(* IEC 61131-3 sources: rusty/tests/lit/single/conversion, 25 files *)

(* ---- to_string_unsupported.st ---- *)
// RUN: not %COMPILE %s 2>&1 | %CHECK %s
// A type with no TO_STRING monomorphization must not silently mis-dispatch to TO_STRING__STRING
// (which reinterprets the argument's bytes and crashes at runtime). Instead the missing
// monomorphization is materialized as an external declaration and surfaces as a link-time undefined
// symbol — a clean, uniform failure for scalar and aggregate returns alike. A user STRUCT never gets
// a monomorph, so this stays valid as follow-up PRs add the remaining scalar conversions.
TYPE MyStruct : STRUCT x : DINT; END_STRUCT END_TYPE

FUNCTION main : DINT
VAR
    st : MyStruct;
    s : STRING;
END_VAR
    // CHECK: {{.*}}TO_STRING__MyStruct{{.*}}
    s := TO_STRING(st);
END_FUNCTION

(* ---- bit_to_real.st ---- *)
// RUN: %COMPILE %s && %RUN | %CHECK %s
//
// BOOL and the bit string types widen to REAL and LREAL by value. BOOL, BYTE and WORD fit a REAL
// exactly, and DWORD fits an LREAL exactly. A REAL keeps 24 bits of mantissa, so a DWORD or LWORD
// above 2^24 is rounded to the nearest representable value on the way in, without a diagnostic.
// These conversions have the named form only; the generic TO_REAL and TO_LREAL take numeric sources.

FUNCTION main
VAR
    umax : LWORD := 0;
END_VAR
umax := umax - 1;   // 2^64 - 1

// BOOL
printf('%.1f %.1f %.1f %.1f$N', BOOL_TO_REAL(FALSE), BOOL_TO_REAL(TRUE), BOOL_TO_LREAL(FALSE), BOOL_TO_LREAL(TRUE));  // CHECK: 0.0 1.0 0.0 1.0

// BYTE and WORD, exact over the whole range
printf('%.0f %.0f %.0f %.0f$N', BYTE_TO_REAL(BYTE#255), BYTE_TO_LREAL(BYTE#255), WORD_TO_REAL(WORD#65535), WORD_TO_LREAL(WORD#65535));  // CHECK: 255 255 65535 65535

// DWORD: exact into LREAL, rounded into REAL above 2^24
printf('%.0f %.0f$N', DWORD_TO_LREAL(DWORD#16777217), DWORD_TO_LREAL(DWORD#4294967295));  // CHECK: 16777217 4294967295
printf('%.0f %.0f$N', DWORD_TO_REAL(DWORD#16777216),  DWORD_TO_REAL(DWORD#16777217));     // CHECK: 16777216 16777216
printf('%.0f$N',      DWORD_TO_REAL(DWORD#4294967295));                                   // CHECK: 4294967296

// LWORD into REAL: 2^24 is the last exact integer
printf('%.0f %.0f$N', LWORD_TO_REAL(LWORD#16777216), LWORD_TO_REAL(LWORD#16777217));          // CHECK: 16777216 16777216
printf('%.0f %.0f$N', LWORD_TO_REAL(LWORD#4294967296), LWORD_TO_REAL(LWORD#9007199254740993));  // CHECK: 4294967296 9007199254740992
printf('%.0f$N',      LWORD_TO_REAL(umax));                                                    // CHECK: 18446744073709551616

// LWORD into LREAL: 2^53 is the last exact integer
printf('%.0f %.0f$N', LWORD_TO_LREAL(LWORD#4611686018427387904), LWORD_TO_LREAL(LWORD#9007199254740993));  // CHECK: 4611686018427387904 9007199254740992
END_FUNCTION

(* ---- num_to_bool.st ---- *)
// RUN: %COMPILE %s && %RUN | %CHECK %s
//
// Every *_TO_BOOL conversion is FALSE for exactly zero and TRUE for everything else. It is not a
// lowest-bit test, a fraction is not truncated first, there is no epsilon, and NaN and the
// infinities are TRUE.

FUNCTION main
VAR
    umax : ULINT := 0;
    ninf : REAL;
END_VAR
umax := umax - 1;   // 2^64 - 1
ninf := -INF_REAL;

// signed integers
printf('%d %d %d %d %d$N', SINT_TO_BOOL(SINT#-128), SINT_TO_BOOL(SINT#0), INT_TO_BOOL(INT#2), INT_TO_BOOL(INT#256), INT_TO_BOOL(INT#-1));  // CHECK: 1 0 1 1 1
printf('%d %d %d %d$N',    INT_TO_BOOL(INT#0), INT_TO_BOOL(INT#1), DINT_TO_BOOL(DINT#65536), LINT_TO_BOOL(LINT#4294967296));                  // CHECK: 0 1 1 1

// unsigned integers
printf('%d %d %d %d$N', USINT_TO_BOOL(USINT#255), USINT_TO_BOOL(USINT#0), UINT_TO_BOOL(UINT#256), UDINT_TO_BOOL(UDINT#4294967295));  // CHECK: 1 0 1 1
printf('%d %d %d %d$N', USINT_TO_BOOL(USINT#1), UINT_TO_BOOL(UINT#0), UINT_TO_BOOL(UINT#65535), UDINT_TO_BOOL(UDINT#65536));         // CHECK: 1 0 1 1
printf('%d %d %d %d$N', ULINT_TO_BOOL(umax), ULINT_TO_BOOL(ULINT#9223372036854775807), ULINT_TO_BOOL(ULINT#4294967296), ULINT_TO_BOOL(ULINT#0));  // CHECK: 1 1 1 0

// reals
printf('%d %d %d %d$N', REAL_TO_BOOL(REAL#0.5), REAL_TO_BOOL(REAL#1.0E-30), REAL_TO_BOOL(REAL#0.0), REAL_TO_BOOL(-REAL#0.0));  // CHECK: 1 1 0 0
printf('%d %d %d$N',    REAL_TO_BOOL(NAN_REAL), REAL_TO_BOOL(INF_REAL), REAL_TO_BOOL(ninf));                                    // CHECK: 1 1 1
printf('%d %d %d$N',    LREAL_TO_BOOL(LREAL#-0.5), LREAL_TO_BOOL(LREAL#0.0), LREAL_TO_BOOL(NAN_LREAL));                          // CHECK: 1 0 1
printf('%d %d %d$N',    LREAL_TO_BOOL(LREAL#0.5), LREAL_TO_BOOL(-LREAL#0.0), LREAL_TO_BOOL(LREAL#1.0E-300));                     // CHECK: 1 0 1

// bit strings, a set bit above bit 0 is TRUE as well
printf('%d %d %d %d %d$N', BYTE_TO_BOOL(BYTE#2), BYTE_TO_BOOL(BYTE#0), WORD_TO_BOOL(WORD#256), DWORD_TO_BOOL(DWORD#65536), LWORD_TO_BOOL(LWORD#4294967296));  // CHECK: 1 0 1 1 1

// the generic form calls the named one
printf('%d %d %d %d$N', TO_BOOL(INT#256), TO_BOOL(REAL#0.5), TO_BOOL(ULINT#4294967296), TO_BOOL(BYTE#2));  // CHECK: 1 1 1 1
END_FUNCTION

(* ---- real_to_bit.st ---- *)
// RUN: %COMPILE %s && %RUN | %CHECK %s
//
// REAL and LREAL to the bit string types round half away from zero, then keep the low bits of the
// target width, so an out-of-range value wraps and a negative value lands at the top of the range.
// The rounded value first becomes a signed 64-bit integer; NaN, the infinities and anything outside
// that range become 2^63 instead, so BYTE, WORD and DWORD see 0 for them. LWORD is the exception:
// a value in [2^63, 2^64) converts exactly, and only NaN, the infinities, values below -2^63 and
// values at or above 2^64 give 2^63. Every cell was measured on CODESYS 3.5 SP22.
FUNCTION main
VAR
    ninf    : REAL;
    lninf   : LREAL;
    band_lo : LREAL := 9223372036854775808.0;   (* 2^63, the smallest LREAL above it is added below *)
    two64   : LREAL := 9223372036854775808.0;
END_VAR
ninf    := -INF_REAL;
lninf   := -INF_LREAL;
band_lo := band_lo + 2048.0;
two64   := two64 * 2.0;

// ---- REAL source: BYTE WORD DWORD LWORD
// rounding, ties away from zero
printf('%d %d %u %llu$N', REAL_TO_BYTE(REAL#0.4),  REAL_TO_WORD(REAL#0.4),  REAL_TO_DWORD(REAL#0.4),  REAL_TO_LWORD(REAL#0.4));   // CHECK: 0 0 0 0
printf('%d %d %u %llu$N', REAL_TO_BYTE(REAL#0.5),  REAL_TO_WORD(REAL#0.5),  REAL_TO_DWORD(REAL#0.5),  REAL_TO_LWORD(REAL#0.5));   // CHECK: 1 1 1 1
printf('%d %d %u %llu$N', REAL_TO_BYTE(REAL#0.6),  REAL_TO_WORD(REAL#0.6),  REAL_TO_DWORD(REAL#0.6),  REAL_TO_LWORD(REAL#0.6));   // CHECK: 1 1 1 1
printf('%d %d %u %llu$N', REAL_TO_BYTE(REAL#1.5),  REAL_TO_WORD(REAL#1.5),  REAL_TO_DWORD(REAL#1.5),  REAL_TO_LWORD(REAL#1.5));   // CHECK: 2 2 2 2
printf('%d %d %u %llu$N', REAL_TO_BYTE(REAL#2.5),  REAL_TO_WORD(REAL#2.5),  REAL_TO_DWORD(REAL#2.5),  REAL_TO_LWORD(REAL#2.5));   // CHECK: 3 3 3 3
printf('%d %d %u %llu$N', REAL_TO_BYTE(REAL#3.5),  REAL_TO_WORD(REAL#3.5),  REAL_TO_DWORD(REAL#3.5),  REAL_TO_LWORD(REAL#3.5));   // CHECK: 4 4 4 4
printf('%d %d %u %llu$N', REAL_TO_BYTE(REAL#-0.5), REAL_TO_WORD(REAL#-0.5), REAL_TO_DWORD(REAL#-0.5), REAL_TO_LWORD(REAL#-0.5));  // CHECK: 255 65535 4294967295 18446744073709551615
printf('%d %d %u %llu$N', REAL_TO_BYTE(REAL#-1.5), REAL_TO_WORD(REAL#-1.5), REAL_TO_DWORD(REAL#-1.5), REAL_TO_LWORD(REAL#-1.5));  // CHECK: 254 65534 4294967294 18446744073709551614
printf('%d %d %u %llu$N', REAL_TO_BYTE(REAL#-2.5), REAL_TO_WORD(REAL#-2.5), REAL_TO_DWORD(REAL#-2.5), REAL_TO_LWORD(REAL#-2.5));  // CHECK: 253 65533 4294967293 18446744073709551613
// range, wraps modulo the target width
printf('%d %d %u %llu$N', REAL_TO_BYTE(REAL#255.5),   REAL_TO_WORD(REAL#255.5),   REAL_TO_DWORD(REAL#255.5),   REAL_TO_LWORD(REAL#255.5));    // CHECK: 0 256 256 256
printf('%d %d %u %llu$N', REAL_TO_BYTE(REAL#256.0),   REAL_TO_WORD(REAL#256.0),   REAL_TO_DWORD(REAL#256.0),   REAL_TO_LWORD(REAL#256.0));    // CHECK: 0 256 256 256
printf('%d %d %u %llu$N', REAL_TO_BYTE(REAL#300.0),   REAL_TO_WORD(REAL#300.0),   REAL_TO_DWORD(REAL#300.0),   REAL_TO_LWORD(REAL#300.0));    // CHECK: 44 300 300 300
printf('%d %d %u %llu$N', REAL_TO_BYTE(REAL#-1.0),    REAL_TO_WORD(REAL#-1.0),    REAL_TO_DWORD(REAL#-1.0),    REAL_TO_LWORD(REAL#-1.0));     // CHECK: 255 65535 4294967295 18446744073709551615
printf('%d %d %u %llu$N', REAL_TO_BYTE(REAL#65536.0), REAL_TO_WORD(REAL#65536.0), REAL_TO_DWORD(REAL#65536.0), REAL_TO_LWORD(REAL#65536.0));  // CHECK: 0 0 65536 65536
printf('%d %d %u %llu$N', REAL_TO_BYTE(REAL#1.0E10),  REAL_TO_WORD(REAL#1.0E10),  REAL_TO_DWORD(REAL#1.0E10),  REAL_TO_LWORD(REAL#1.0E10));   // CHECK: 0 58368 1410065408 10000000000
printf('%d %d %u %llu$N', REAL_TO_BYTE(REAL#1.0E20),  REAL_TO_WORD(REAL#1.0E20),  REAL_TO_DWORD(REAL#1.0E20),  REAL_TO_LWORD(REAL#1.0E20));   // CHECK: 0 0 0 9223372036854775808
// not a number
printf('%d %d %u %llu$N', REAL_TO_BYTE(INF_REAL), REAL_TO_WORD(INF_REAL), REAL_TO_DWORD(INF_REAL), REAL_TO_LWORD(INF_REAL));  // CHECK: 0 0 0 9223372036854775808
printf('%d %d %u %llu$N', REAL_TO_BYTE(ninf),     REAL_TO_WORD(ninf),     REAL_TO_DWORD(ninf),     REAL_TO_LWORD(ninf));      // CHECK: 0 0 0 9223372036854775808
printf('%d %d %u %llu$N', REAL_TO_BYTE(NAN_REAL), REAL_TO_WORD(NAN_REAL), REAL_TO_DWORD(NAN_REAL), REAL_TO_LWORD(NAN_REAL));  // CHECK: 0 0 0 9223372036854775808

// ---- LREAL source: BYTE WORD DWORD LWORD
printf('%d %d %u %llu$N', LREAL_TO_BYTE(LREAL#0.5),     LREAL_TO_WORD(LREAL#0.5),     LREAL_TO_DWORD(LREAL#0.5),     LREAL_TO_LWORD(LREAL#0.5));      // CHECK: 1 1 1 1
printf('%d %d %u %llu$N', LREAL_TO_BYTE(LREAL#2.5),     LREAL_TO_WORD(LREAL#2.5),     LREAL_TO_DWORD(LREAL#2.5),     LREAL_TO_LWORD(LREAL#2.5));      // CHECK: 3 3 3 3
printf('%d %d %u %llu$N', LREAL_TO_BYTE(LREAL#-0.5),    LREAL_TO_WORD(LREAL#-0.5),    LREAL_TO_DWORD(LREAL#-0.5),    LREAL_TO_LWORD(LREAL#-0.5));     // CHECK: 255 65535 4294967295 18446744073709551615
printf('%d %d %u %llu$N', LREAL_TO_BYTE(LREAL#-2.5),    LREAL_TO_WORD(LREAL#-2.5),    LREAL_TO_DWORD(LREAL#-2.5),    LREAL_TO_LWORD(LREAL#-2.5));     // CHECK: 253 65533 4294967293 18446744073709551613
printf('%d %d %u %llu$N', LREAL_TO_BYTE(LREAL#255.5),   LREAL_TO_WORD(LREAL#255.5),   LREAL_TO_DWORD(LREAL#255.5),   LREAL_TO_LWORD(LREAL#255.5));    // CHECK: 0 256 256 256
printf('%d %d %u %llu$N', LREAL_TO_BYTE(LREAL#300.0),   LREAL_TO_WORD(LREAL#300.0),   LREAL_TO_DWORD(LREAL#300.0),   LREAL_TO_LWORD(LREAL#300.0));    // CHECK: 44 300 300 300
printf('%d %d %u %llu$N', LREAL_TO_BYTE(LREAL#-1.0),    LREAL_TO_WORD(LREAL#-1.0),    LREAL_TO_DWORD(LREAL#-1.0),    LREAL_TO_LWORD(LREAL#-1.0));     // CHECK: 255 65535 4294967295 18446744073709551615
printf('%d %d %u %llu$N', LREAL_TO_BYTE(LREAL#65536.0), LREAL_TO_WORD(LREAL#65536.0), LREAL_TO_DWORD(LREAL#65536.0), LREAL_TO_LWORD(LREAL#65536.0));  // CHECK: 0 0 65536 65536
printf('%d %d %u %llu$N', LREAL_TO_BYTE(LREAL#1.0E10),  LREAL_TO_WORD(LREAL#1.0E10),  LREAL_TO_DWORD(LREAL#1.0E10),  LREAL_TO_LWORD(LREAL#1.0E10));   // CHECK: 0 58368 1410065408 10000000000
printf('%d %d %u %llu$N', LREAL_TO_BYTE(LREAL#1.0E20),  LREAL_TO_WORD(LREAL#1.0E20),  LREAL_TO_DWORD(LREAL#1.0E20),  LREAL_TO_LWORD(LREAL#1.0E20));   // CHECK: 0 0 0 9223372036854775808
printf('%d %d %u %llu$N', LREAL_TO_BYTE(INF_LREAL), LREAL_TO_WORD(INF_LREAL), LREAL_TO_DWORD(INF_LREAL), LREAL_TO_LWORD(INF_LREAL));  // CHECK: 0 0 0 9223372036854775808
printf('%d %d %u %llu$N', LREAL_TO_BYTE(lninf),     LREAL_TO_WORD(lninf),     LREAL_TO_DWORD(lninf),     LREAL_TO_LWORD(lninf));      // CHECK: 0 0 0 9223372036854775808
printf('%d %d %u %llu$N', LREAL_TO_BYTE(NAN_LREAL), LREAL_TO_WORD(NAN_LREAL), LREAL_TO_DWORD(NAN_LREAL), LREAL_TO_LWORD(NAN_LREAL));  // CHECK: 0 0 0 9223372036854775808

// ---- the 64-bit band: LWORD keeps [2^63, 2^64) exact, the narrower targets go through the signed path
printf('%u %llu$N', LREAL_TO_DWORD(LREAL#1.0E19), LREAL_TO_LWORD(LREAL#1.0E19));   // CHECK: 0 10000000000000000000
printf('%llu %llu$N', LREAL_TO_LWORD(band_lo), LREAL_TO_LWORD(LREAL#1.8E19));      // CHECK: 9223372036854777856 18000000000000000000
printf('%llu %llu$N', LREAL_TO_LWORD(two64), LREAL_TO_LWORD(LREAL#-1.0E19));       // CHECK: 9223372036854775808 9223372036854775808
printf('%llu$N', REAL_TO_LWORD(REAL#1.0E19));                                       // CHECK: 9999999980506447872

// ---- the generic form calls the named one
printf('%d %d %u %llu$N', TO_BYTE(REAL#300.0), TO_WORD(LREAL#-1.0), TO_DWORD(REAL#1.0E10), TO_LWORD(LREAL#-0.5));  // CHECK: 44 65535 1410065408 18446744073709551615
END_FUNCTION

(* ---- real_trunc_int.st ---- *)
// RUN: %COMPILE %s && %RUN | %CHECK %s
FUNCTION main
    printf('%d$N', REAL_TRUNC_SINT(5.6));       // CHECK: 5
    printf('%d$N', REAL_TRUNC_USINT(5.6));      // CHECK: 5
    printf('%d$N', REAL_TRUNC_INT(5.6));        // CHECK: 5
    printf('%d$N', REAL_TRUNC_UINT(5.6));       // CHECK: 5
    printf('%d$N', REAL_TRUNC_INT(5.6));        // CHECK: 5
    printf('%d$N', REAL_TRUNC_UINT(5.6));       // CHECK: 5
    printf('%d$N', REAL_TRUNC_DINT(5.6));       // CHECK: 5
    printf('%d$N', REAL_TRUNC_UDINT(5.6));      // CHECK: 5
    printf('%d$N', REAL_TRUNC_LINT(5.6));       // CHECK: 5
    printf('%d$N', REAL_TRUNC_ULINT(5.6));      // CHECK: 5

    printf('%d$N', REAL_TRUNC_SINT(-5.6));      // CHECK: -5
    printf('%d$N', REAL_TRUNC_INT(-5.6));       // CHECK: -5
    printf('%d$N', REAL_TRUNC_DINT(-5.6));      // CHECK: -5
    printf('%d$N', REAL_TRUNC_LINT(-5.6));      // CHECK: -5
END_FUNCTION

(* ---- string_to_based_literals.st ---- *)
// STRING_TO integer and bit-string conversions accept IEC based literals and nothing else.
// RUN: %COMPILE %s && %RUN | %CHECK %s

FUNCTION main
    printf('byte_hex=%d$N', STRING_TO_BYTE('16#FF'));        // CHECK: byte_hex=255
    printf('word_octal=%d$N', STRING_TO_WORD('8#777'));      // CHECK-NEXT: word_octal=511
    printf('dword_binary=%d$N', STRING_TO_DWORD('2#1010'));  // CHECK-NEXT: dword_binary=10
    printf('dint_binary=%d$N', STRING_TO_DINT('2#1010'));    // CHECK-NEXT: dint_binary=10
    printf('lint_binary=%d$N', STRING_TO_LINT('2#1010'));    // CHECK-NEXT: lint_binary=10
    printf('lword_lower_hex=%d$N', STRING_TO_LWORD('16#ff'));// CHECK-NEXT: lword_lower_hex=255
    printf('dint_hex=%d$N', STRING_TO_DINT('16#FF'));        // CHECK-NEXT: dint_hex=255
    printf('lint_hex=%d$N', STRING_TO_LINT('16#FF'));        // CHECK-NEXT: lint_hex=255
    printf('dint_octal=%d$N', STRING_TO_DINT('8#77'));       // CHECK-NEXT: dint_octal=63
    printf('lint_octal=%d$N', STRING_TO_LINT('8#77'));       // CHECK-NEXT: lint_octal=63
    printf('udint_grouped_hex=%d$N', STRING_TO_UDINT('16#FF_FF')); // CHECK-NEXT: udint_grouped_hex=65535
    printf('ulint_trimmed_hex=%d$N', STRING_TO_ULINT(' 16#FF ')); // CHECK-NEXT: ulint_trimmed_hex=255
    printf('missing_digits=%d$N', STRING_TO_UDINT('16#'));   // CHECK-NEXT: missing_digits=0
    printf('invalid_digit=%d$N', STRING_TO_UDINT('16#GG'));  // CHECK-NEXT: invalid_digit=0
    printf('unsupported_radix=%d$N', STRING_TO_UDINT('10#42')); // CHECK-NEXT: unsupported_radix=0
    printf('signed_hex=%d$N', STRING_TO_UDINT('+16#FF'));    // CHECK-NEXT: signed_hex=0

    // Based literals are unsigned; a sign on either side of the radix is rejected.
    printf('negative_hex=%d$N', STRING_TO_DINT('-16#FF'));   // CHECK-NEXT: negative_hex=0
    printf('hex_negative=%d$N', STRING_TO_DINT('16#-FF'));   // CHECK-NEXT: hex_negative=0
    printf('binary_negative=%d$N', STRING_TO_SINT('2#-1'));  // CHECK-NEXT: binary_negative=0

    // Underscores group digits; they may not lead, trail or double up.
    printf('leading_underscore=%d$N', STRING_TO_UDINT('16#_FF'));  // CHECK-NEXT: leading_underscore=0
    printf('trailing_underscore=%d$N', STRING_TO_UDINT('16#FF_')); // CHECK-NEXT: trailing_underscore=0
    printf('double_underscore=%d$N', STRING_TO_UDINT('16#F__F')); // CHECK-NEXT: double_underscore=0
    printf('decimal_grouped=%d$N', STRING_TO_UDINT('1_000'));     // CHECK-NEXT: decimal_grouped=1000
    printf('decimal_leading_us=%d$N', STRING_TO_UDINT('_1'));     // CHECK-NEXT: decimal_leading_us=0
    printf('decimal_double_us=%d$N', STRING_TO_UDINT('1__0'));    // CHECK-NEXT: decimal_double_us=0

    // C-style radix prefixes are not Structured Text literals.
    printf('byte_c_binary=%d$N', STRING_TO_BYTE('0b1010'));   // CHECK-NEXT: byte_c_binary=0
    printf('lword_c_binary=%d$N', STRING_TO_LWORD('0B1010')); // CHECK-NEXT: lword_c_binary=0
    printf('dint_c_hex=%d$N', STRING_TO_DINT('0x7F'));        // CHECK-NEXT: dint_c_hex=0
    printf('ulint_c_hex=%d$N', STRING_TO_ULINT('0X7F'));      // CHECK-NEXT: ulint_c_hex=0

    // A hexadecimal bit pattern that does not fit the signed target is rejected, not reinterpreted.
    printf('int_hex_max=%d$N', STRING_TO_INT('16#7FFF'));          // CHECK-NEXT: int_hex_max=32767
    printf('int_hex_all_ones=%d$N', STRING_TO_INT('16#FFFF'));     // CHECK-NEXT: int_hex_all_ones=0
    printf('word_hex_all_ones=%d$N', STRING_TO_WORD('16#FFFF'));   // CHECK-NEXT: word_hex_all_ones=65535
END_FUNCTION

(* ---- string_to_bool.st ---- *)
// STRING_TO_BOOL accepts true values and rejects malformed values.
// RUN: %COMPILE %s && %RUN | %CHECK %s

FUNCTION main
    printf('garbage=%d$N', STRING_TO_BOOL('garbage'));       // CHECK: garbage=0
    printf('numeric_one=%d$N', STRING_TO_BOOL('1'));         // CHECK-NEXT: numeric_one=1
    printf('upper_true=%d$N', STRING_TO_BOOL('TRUE'));       // CHECK-NEXT: upper_true=1
    printf('lower_true=%d$N', STRING_TO_BOOL('true'));       // CHECK-NEXT: lower_true=1
    printf('trimmed_true=%d$N', STRING_TO_BOOL('  true  ')); // CHECK-NEXT: trimmed_true=1
    printf('numeric_zero=%d$N', STRING_TO_BOOL('0'));        // CHECK-NEXT: numeric_zero=0
    printf('numeric_two=%d$N', STRING_TO_BOOL('2'));         // CHECK-NEXT: numeric_two=0
    printf('false=%d$N', STRING_TO_BOOL('false'));           // CHECK-NEXT: false=0
    printf('suffix=%d$N', STRING_TO_BOOL('TRUEX'));          // CHECK-NEXT: suffix=0
END_FUNCTION

(* ---- string_to_calendar.st ---- *)
// STRING_TO_DATE, STRING_TO_DT, and STRING_TO_TOD accept exactly the calendar literals of their type.
// RUN: %COMPILE %s && %RUN | %CHECK %s

FUNCTION main
    // Valid prefixed literals parse for each target type.
    printf('date_valid=%s$N', REF(DATE_TO_STRING(STRING_TO_DATE('D#2024-02-29')))); // CHECK: date_valid=D#2024-02-29
    printf('dt_valid=%s$N', REF(DT_TO_STRING(STRING_TO_DT('DT#2024-01-01-12:00:00')))); // CHECK-NEXT: dt_valid=DT#2024-01-01-12:00:00
    printf('tod_valid=%s$N', REF(TOD_TO_STRING(STRING_TO_TOD('TOD#12:00:00')))); // CHECK-NEXT: tod_valid=TOD#12:00:00

    // Empty input returns each type's zero value.
    printf('date_empty=%s$N', REF(DATE_TO_STRING(STRING_TO_DATE('')))); // CHECK-NEXT: date_empty=D#1970-01-01
    printf('dt_empty=%s$N', REF(DT_TO_STRING(STRING_TO_DT('')))); // CHECK-NEXT: dt_empty=DT#1970-01-01-00:00:00
    printf('tod_empty=%s$N', REF(TOD_TO_STRING(STRING_TO_TOD('')))); // CHECK-NEXT: tod_empty=TOD#00:00:00

    // Malformed input returns each type's zero value.
    printf('date_garbage=%s$N', REF(DATE_TO_STRING(STRING_TO_DATE('not a date')))); // CHECK-NEXT: date_garbage=D#1970-01-01
    printf('dt_garbage=%s$N', REF(DT_TO_STRING(STRING_TO_DT('$00')))); // CHECK-NEXT: dt_garbage=DT#1970-01-01-00:00:00
    printf('tod_garbage=%s$N', REF(TOD_TO_STRING(STRING_TO_TOD('bad')))); // CHECK-NEXT: tod_garbage=TOD#00:00:00

    // Each conversion rejects a literal prefix for a different calendar type.
    printf('date_wrong_prefix=%s$N', REF(DATE_TO_STRING(STRING_TO_DATE('TOD#12:45:00')))); // CHECK-NEXT: date_wrong_prefix=D#1970-01-01
    printf('dt_wrong_prefix=%s$N', REF(DT_TO_STRING(STRING_TO_DT('D#2024-01-01')))); // CHECK-NEXT: dt_wrong_prefix=DT#1970-01-01-00:00:00
    printf('tod_wrong_prefix=%s$N', REF(TOD_TO_STRING(STRING_TO_TOD('DT#2024-01-01-12:00:00')))); // CHECK-NEXT: tod_wrong_prefix=TOD#00:00:00

    // Out-of-range date and time fields are rejected.
    printf('date_invalid_day=%s$N', REF(DATE_TO_STRING(STRING_TO_DATE('D#2024-02-30')))); // CHECK-NEXT: date_invalid_day=D#1970-01-01
    printf('dt_invalid_hour=%s$N', REF(DT_TO_STRING(STRING_TO_DT('DT#2024-01-01-25:00:00')))); // CHECK-NEXT: dt_invalid_hour=DT#1970-01-01-00:00:00
    printf('tod_invalid_minute=%s$N', REF(TOD_TO_STRING(STRING_TO_TOD('TOD#12:60:00')))); // CHECK-NEXT: tod_invalid_minute=TOD#00:00:00

    // Values outside the representable range return the zero value.
    printf('date_low_range=%s$N', REF(DATE_TO_STRING(STRING_TO_DATE('D#1969-12-31')))); // CHECK-NEXT: date_low_range=D#1970-01-01
    printf('dt_low_range=%s$N', REF(DT_TO_STRING(STRING_TO_DT('DT#1969-12-31-23:59:59')))); // CHECK-NEXT: dt_low_range=DT#1970-01-01-00:00:00
    printf('tod_high_range=%s$N', REF(TOD_TO_STRING(STRING_TO_TOD('TOD#25:00:00')))); // CHECK-NEXT: tod_high_range=TOD#00:00:00
    printf('date_high_range=%s$N', REF(DATE_TO_STRING(STRING_TO_DATE('D#2106-02-08')))); // CHECK-NEXT: date_high_range=D#1970-01-01
    printf('dt_high_range=%s$N', REF(DT_TO_STRING(STRING_TO_DT('DT#2106-02-08-00:00:00')))); // CHECK-NEXT: dt_high_range=DT#1970-01-01-00:00:00
    printf('tod_low_range=%s$N', REF(TOD_TO_STRING(STRING_TO_TOD('TOD#-1:00:00')))); // CHECK-NEXT: tod_low_range=TOD#00:00:00

    // DATE rejects fractions, DT drops them, and TOD preserves milliseconds.
    printf('date_fraction=%s$N', REF(DATE_TO_STRING(STRING_TO_DATE('D#2024-01-01.500')))); // CHECK-NEXT: date_fraction=D#1970-01-01
    printf('dt_fraction=%s$N', REF(DT_TO_STRING(STRING_TO_DT('DT#2024-01-01-12:00:00.500')))); // CHECK-NEXT: dt_fraction=DT#2024-01-01-12:00:00
    printf('tod_fraction=%s$N', REF(TOD_TO_STRING(STRING_TO_TOD('TOD#12:00:00.500')))); // CHECK-NEXT: tod_fraction=TOD#12:00:00.500

    // The literal prefix is required; bare ISO forms are rejected.
    printf('date_unprefixed=%s$N', REF(DATE_TO_STRING(STRING_TO_DATE('2024-01-01')))); // CHECK-NEXT: date_unprefixed=D#1970-01-01
    printf('dt_unprefixed_date=%s$N', REF(DT_TO_STRING(STRING_TO_DT('2024-01-01')))); // CHECK-NEXT: dt_unprefixed_date=DT#1970-01-01-00:00:00
    printf('dt_unprefixed=%s$N', REF(DT_TO_STRING(STRING_TO_DT('2024-01-01T12:00:00')))); // CHECK-NEXT: dt_unprefixed=DT#1970-01-01-00:00:00
    printf('tod_unprefixed=%s$N', REF(TOD_TO_STRING(STRING_TO_TOD('12:00:00')))); // CHECK-NEXT: tod_unprefixed=TOD#00:00:00

    // The long spelling of each prefix is accepted, case-insensitively.
    printf('date_long_prefix=%s$N', REF(DATE_TO_STRING(STRING_TO_DATE('date#2024-01-01')))); // CHECK-NEXT: date_long_prefix=D#2024-01-01
    printf('dt_long_prefix=%s$N', REF(DT_TO_STRING(STRING_TO_DT('DATE_AND_TIME#2024-01-01-12:00:00')))); // CHECK-NEXT: dt_long_prefix=DT#2024-01-01-12:00:00
    printf('tod_long_prefix=%s$N', REF(TOD_TO_STRING(STRING_TO_TOD('time_of_day#12:00:00')))); // CHECK-NEXT: tod_long_prefix=TOD#12:00:00

    // The 64-bit literal prefixes belong to LDATE, LDT and LTOD and are rejected here.
    printf('date_ldate_prefix=%s$N', REF(DATE_TO_STRING(STRING_TO_DATE('LDATE#2024-01-01')))); // CHECK-NEXT: date_ldate_prefix=D#1970-01-01
    printf('dt_ldt_prefix=%s$N', REF(DT_TO_STRING(STRING_TO_DT('LDT#2024-01-01-12:00:00')))); // CHECK-NEXT: dt_ldt_prefix=DT#1970-01-01-00:00:00
    printf('tod_ltod_prefix=%s$N', REF(TOD_TO_STRING(STRING_TO_TOD('LTOD#12:00:00')))); // CHECK-NEXT: tod_ltod_prefix=TOD#00:00:00

    // Nothing may follow the literal, not even comment-like text.
    printf('date_trailing=%s$N', REF(DATE_TO_STRING(STRING_TO_DATE('D#2024-01-01//x')))); // CHECK-NEXT: date_trailing=D#1970-01-01
    printf('dt_trailing=%s$N', REF(DT_TO_STRING(STRING_TO_DT('DT#2024-01-01-12:00:00(*x*)')))); // CHECK-NEXT: dt_trailing=DT#1970-01-01-00:00:00
    printf('tod_trailing=%s$N', REF(TOD_TO_STRING(STRING_TO_TOD('TOD#12:00:00{x}')))); // CHECK-NEXT: tod_trailing=TOD#00:00:00

    // Fractions truncate: no rounding into the next second or day.
    printf('tod_truncated=%s$N', REF(TOD_TO_STRING(STRING_TO_TOD('TOD#23:59:59.9999999999')))); // CHECK-NEXT: tod_truncated=TOD#23:59:59.999
    printf('dt_truncated=%s$N', REF(DT_TO_STRING(STRING_TO_DT('DT#2024-01-01-23:59:59.9999999999')))); // CHECK-NEXT: dt_truncated=DT#2024-01-01-23:59:59

    // Single-digit fields and optional seconds follow the literal grammar.
    printf('date_short_fields=%s$N', REF(DATE_TO_STRING(STRING_TO_DATE('D#2024-1-1')))); // CHECK-NEXT: date_short_fields=D#2024-01-01
    printf('dt_no_seconds=%s$N', REF(DT_TO_STRING(STRING_TO_DT('DT#2024-01-01-12:00')))); // CHECK-NEXT: dt_no_seconds=DT#2024-01-01-12:00:00
    printf('tod_no_seconds=%s$N', REF(TOD_TO_STRING(STRING_TO_TOD('TOD#12:00')))); // CHECK-NEXT: tod_no_seconds=TOD#12:00:00

    // Surrounding whitespace is ignored for every target type.
    printf('date_trimmed=%s$N', REF(DATE_TO_STRING(STRING_TO_DATE(' D#2024-01-01 ')))); // CHECK-NEXT: date_trimmed=D#2024-01-01
    printf('dt_trimmed=%s$N', REF(DT_TO_STRING(STRING_TO_DT('$TDT#2024-01-01-12:00:00$R$N')))); // CHECK-NEXT: dt_trimmed=DT#2024-01-01-12:00:00
    printf('tod_trimmed=%s$N', REF(TOD_TO_STRING(STRING_TO_TOD('$TTOD#12:00:00$T')))); // CHECK-NEXT: tod_trimmed=TOD#12:00:00

    // Whitespace within a literal is rejected for every target type.
    printf('date_internal_space=%s$N', REF(DATE_TO_STRING(STRING_TO_DATE('D# 2024-01-01')))); // CHECK-NEXT: date_internal_space=D#1970-01-01
    printf('dt_internal_space=%s$N', REF(DT_TO_STRING(STRING_TO_DT('DT#2024-01-01 12:00:00')))); // CHECK-NEXT: dt_internal_space=DT#1970-01-01-00:00:00
    printf('tod_internal_space=%s$N', REF(TOD_TO_STRING(STRING_TO_TOD('TOD#12: 00:00')))); // CHECK-NEXT: tod_internal_space=TOD#00:00:00
END_FUNCTION

(* ---- string_to_duration.st ---- *)
// STRING_TO_TIME and STRING_TO_LTIME parse duration literals with exact arithmetic.
// RUN: %COMPILE %s && %RUN | %CHECK %s

FUNCTION main
    printf('time_fraction_1_5s=%s$N', REF(TIME_TO_STRING(STRING_TO_TIME('T#1.5s')))); // CHECK: time_fraction_1_5s=T#1s500ms
    printf('time_fraction_0_5s=%s$N', REF(TIME_TO_STRING(STRING_TO_TIME('T#0.5s')))); // CHECK-NEXT: time_fraction_0_5s=T#500ms
    printf('time_fraction_2_75s=%s$N', REF(TIME_TO_STRING(STRING_TO_TIME('T#2.75s')))); // CHECK-NEXT: time_fraction_2_75s=T#2s750ms
    printf('time_fraction_comma=%s$N', REF(TIME_TO_STRING(STRING_TO_TIME('T#1,5s')))); // CHECK-NEXT: time_fraction_comma=T#0ms
    printf('time_fraction_inner=%s$N', REF(TIME_TO_STRING(STRING_TO_TIME('T#1.5h30m')))); // CHECK-NEXT: time_fraction_inner=T#2h
    printf('time_fraction_resolution=%s$N', REF(TIME_TO_STRING(STRING_TO_TIME('T#1.0004ms')))); // CHECK-NEXT: time_fraction_resolution=T#1ms
    printf('ltime_fraction=%s$N', REF(LTIME_TO_STRING(STRING_TO_LTIME('LTIME#1.5s')))); // CHECK-NEXT: ltime_fraction=LTIME#1s500ms
    printf('time_compound=%s$N', REF(TIME_TO_STRING(STRING_TO_TIME('TIME#1d2h3m4s5ms')))); // CHECK-NEXT: time_compound=T#1d2h3m4s5ms
    printf('time_case_insensitive=%s$N', REF(TIME_TO_STRING(STRING_TO_TIME('time#1s')))); // CHECK-NEXT: time_case_insensitive=T#1s
    printf('ltime_nanoseconds=%s$N', REF(LTIME_TO_STRING(STRING_TO_LTIME('LT#1ns')))); // CHECK-NEXT: ltime_nanoseconds=LTIME#1ns
    printf('time_negative=%s$N', REF(TIME_TO_STRING(STRING_TO_TIME('T#-1s')))); // CHECK-NEXT: time_negative=T#0ms
    printf('ltime_negative=%s$N', REF(LTIME_TO_STRING(STRING_TO_LTIME('LTIME#-1s')))); // CHECK-NEXT: ltime_negative=LTIME#0ns
    printf('time_empty=%s$N', REF(TIME_TO_STRING(STRING_TO_TIME('')))); // CHECK-NEXT: time_empty=T#0ms
    printf('time_garbage=%s$N', REF(TIME_TO_STRING(STRING_TO_TIME('abc')))); // CHECK-NEXT: time_garbage=T#0ms
    printf('time_missing_prefix=%s$N', REF(TIME_TO_STRING(STRING_TO_TIME('1s')))); // CHECK-NEXT: time_missing_prefix=T#0ms
    printf('time_wrong_prefix=%s$N', REF(TIME_TO_STRING(STRING_TO_TIME('LTIME#1s')))); // CHECK-NEXT: time_wrong_prefix=T#0ms
    printf('time_wrong_formatter=%s$N', REF(TIME_TO_STRING(STRING_TO_TIME('TOD#12:45:00')))); // CHECK-NEXT: time_wrong_formatter=T#0ms
    printf('time_67ms=%s$N', REF(TIME_TO_STRING(STRING_TO_TIME('T#67ms')))); // CHECK-NEXT: time_67ms=T#67ms
    printf('ltime_wrong_formatter=%s$N', REF(LTIME_TO_STRING(STRING_TO_LTIME('T#1s')))); // CHECK-NEXT: ltime_wrong_formatter=LTIME#0ns
    printf('time_missing_unit=%s$N', REF(TIME_TO_STRING(STRING_TO_TIME('T#1000')))); // CHECK-NEXT: time_missing_unit=T#0ms
    printf('time_internal_space=%s$N', REF(TIME_TO_STRING(STRING_TO_TIME('T#1h 30m')))); // CHECK-NEXT: time_internal_space=T#1h30m
    printf('time_underscore_separator=%s$N', REF(TIME_TO_STRING(STRING_TO_TIME('T#1h_30m')))); // CHECK-NEXT: time_underscore_separator=T#1h30m
    printf('time_split_number=%s$N', REF(TIME_TO_STRING(STRING_TO_TIME('T#1 0s')))); // CHECK-NEXT: time_split_number=T#0ms
    printf('time_unordered=%s$N', REF(TIME_TO_STRING(STRING_TO_TIME('T#30m1h')))); // CHECK-NEXT: time_unordered=T#1h30m
    printf('time_repeated=%s$N', REF(TIME_TO_STRING(STRING_TO_TIME('T#1h1h')))); // CHECK-NEXT: time_repeated=T#2h
    printf('time_plus=%s$N', REF(TIME_TO_STRING(STRING_TO_TIME('T#+1s')))); // CHECK-NEXT: time_plus=T#1s
    printf('time_digit_group=%s$N', REF(TIME_TO_STRING(STRING_TO_TIME('T#1_000ms')))); // CHECK-NEXT: time_digit_group=T#1s
    printf('time_trailing=%s$N', REF(TIME_TO_STRING(STRING_TO_TIME('T#1h§30m')))); // CHECK-NEXT: time_trailing=T#0ms
    printf('time_trailing_comment=%s$N', REF(TIME_TO_STRING(STRING_TO_TIME('T#1s//x')))); // CHECK-NEXT: time_trailing_comment=T#0ms
    printf('time_big_ns=%s$N', REF(TIME_TO_STRING(STRING_TO_TIME('T#5000000000ns')))); // CHECK-NEXT: time_big_ns=T#5s
    printf('time_max=%s$N', REF(TIME_TO_STRING(STRING_TO_TIME('T#49d17h2m47s295ms')))); // CHECK-NEXT: time_max=T#49d17h2m47s295ms
    printf('time_overflow=%s$N', REF(TIME_TO_STRING(STRING_TO_TIME('T#49d17h2m47s296ms')))); // CHECK-NEXT: time_overflow=T#0ms
    printf('ltime_max=%s$N', REF(LTIME_TO_STRING(STRING_TO_LTIME('LTIME#106751d23h47m16s854ms775us807ns')))); // CHECK-NEXT: ltime_max=LTIME#106751d23h47m16s854ms775us807ns
    printf('ltime_overflow=%s$N', REF(LTIME_TO_STRING(STRING_TO_LTIME('LTIME#106751d23h47m16s854ms775us808ns')))); // CHECK-NEXT: ltime_overflow=LTIME#0ns
END_FUNCTION

(* ---- string_to_integer.st ---- *)
// STRING_TO integer and bit-string conversions share one parser at every width.
// RUN: %COMPILE %s && %RUN | %CHECK %s

FUNCTION main
    // Empty input returns zero for every target type.
    printf('byte_empty=%d$N', STRING_TO_BYTE(''));       // CHECK: byte_empty=0
    printf('word_empty=%d$N', STRING_TO_WORD(''));       // CHECK-NEXT: word_empty=0
    printf('dword_empty=%d$N', STRING_TO_DWORD(''));     // CHECK-NEXT: dword_empty=0
    printf('lword_empty=%d$N', STRING_TO_LWORD(''));     // CHECK-NEXT: lword_empty=0
    printf('sint_empty=%d$N', STRING_TO_SINT(''));       // CHECK-NEXT: sint_empty=0
    printf('usint_empty=%d$N', STRING_TO_USINT(''));     // CHECK-NEXT: usint_empty=0
    printf('int_empty=%d$N', STRING_TO_INT(''));         // CHECK-NEXT: int_empty=0
    printf('uint_empty=%d$N', STRING_TO_UINT(''));       // CHECK-NEXT: uint_empty=0
    printf('dint_empty=%d$N', STRING_TO_DINT(''));       // CHECK-NEXT: dint_empty=0
    printf('udint_empty=%d$N', STRING_TO_UDINT(''));     // CHECK-NEXT: udint_empty=0
    printf('lint_empty=%d$N', STRING_TO_LINT(''));       // CHECK-NEXT: lint_empty=0
    printf('ulint_empty=%d$N', STRING_TO_ULINT(''));     // CHECK-NEXT: ulint_empty=0

    // Negative input is preserved by signed targets and rejected by unsigned targets.
    printf('byte_negative=%d$N', STRING_TO_BYTE('-1'));  // CHECK-NEXT: byte_negative=0
    printf('word_negative=%d$N', STRING_TO_WORD('-1'));  // CHECK-NEXT: word_negative=0
    printf('dword_negative=%d$N', STRING_TO_DWORD('-1'));// CHECK-NEXT: dword_negative=0
    printf('lword_negative=%d$N', STRING_TO_LWORD('-1'));// CHECK-NEXT: lword_negative=0
    printf('sint_negative=%d$N', STRING_TO_SINT('-1'));  // CHECK-NEXT: sint_negative=-1
    printf('usint_negative=%d$N', STRING_TO_USINT('-1'));// CHECK-NEXT: usint_negative=0
    printf('int_negative=%d$N', STRING_TO_INT('-1'));    // CHECK-NEXT: int_negative=-1
    printf('uint_negative=%d$N', STRING_TO_UINT('-1'));  // CHECK-NEXT: uint_negative=0
    printf('dint_negative=%d$N', STRING_TO_DINT('-1'));  // CHECK-NEXT: dint_negative=-1
    printf('udint_negative=%d$N', STRING_TO_UDINT('-1'));// CHECK-NEXT: udint_negative=0
    printf('lint_negative=%d$N', STRING_TO_LINT('-1'));  // CHECK-NEXT: lint_negative=-1
    printf('ulint_negative=%d$N', STRING_TO_ULINT('-1'));// CHECK-NEXT: ulint_negative=0

    // Malformed input returns zero for every target type.
    printf('byte_malformed=%d$N', STRING_TO_BYTE('12abc'));   // CHECK-NEXT: byte_malformed=0
    printf('word_malformed=%d$N', STRING_TO_WORD('12abc'));   // CHECK-NEXT: word_malformed=0
    printf('dword_malformed=%d$N', STRING_TO_DWORD('12abc')); // CHECK-NEXT: dword_malformed=0
    printf('lword_malformed=%d$N', STRING_TO_LWORD('12abc')); // CHECK-NEXT: lword_malformed=0
    printf('sint_malformed=%d$N', STRING_TO_SINT('12abc'));   // CHECK-NEXT: sint_malformed=0
    printf('usint_malformed=%d$N', STRING_TO_USINT('12abc')); // CHECK-NEXT: usint_malformed=0
    printf('int_malformed=%d$N', STRING_TO_INT('12abc'));     // CHECK-NEXT: int_malformed=0
    printf('uint_malformed=%d$N', STRING_TO_UINT('12abc'));   // CHECK-NEXT: uint_malformed=0
    printf('dint_malformed=%d$N', STRING_TO_DINT('12abc'));   // CHECK-NEXT: dint_malformed=0
    printf('udint_malformed=%d$N', STRING_TO_UDINT('12abc')); // CHECK-NEXT: udint_malformed=0
    printf('lint_malformed=%d$N', STRING_TO_LINT('12abc'));   // CHECK-NEXT: lint_malformed=0
    printf('ulint_malformed=%d$N', STRING_TO_ULINT('12abc')); // CHECK-NEXT: ulint_malformed=0

    // Values that do not fit the target yield zero instead of wrapping.
    printf('byte_overflow=%d$N', STRING_TO_BYTE('256'));                   // CHECK-NEXT: byte_overflow=0
    printf('sint_overflow=%d$N', STRING_TO_SINT('128'));                   // CHECK-NEXT: sint_overflow=0
    printf('int_overflow=%d$N', STRING_TO_INT('32768'));                   // CHECK-NEXT: int_overflow=0
    printf('dint_overflow=%d$N', STRING_TO_DINT('2147483648'));            // CHECK-NEXT: dint_overflow=0
    printf('dint_underflow=%d$N', STRING_TO_DINT('-2147483649'));          // CHECK-NEXT: dint_underflow=0
    printf('udint_overflow=%d$N', STRING_TO_UDINT('4294967296'));          // CHECK-NEXT: udint_overflow=0
    printf('lint_overflow=%d$N', STRING_TO_LINT('9223372036854775808'));   // CHECK-NEXT: lint_overflow=0
    printf('ulint_overflow=%d$N', STRING_TO_ULINT('18446744073709551616'));// CHECK-NEXT: ulint_overflow=0
    printf('dint_max=%d$N', STRING_TO_DINT('2147483647'));                 // CHECK-NEXT: dint_max=2147483647
    printf('dint_min=%d$N', STRING_TO_DINT('-2147483648'));                // CHECK-NEXT: dint_min=-2147483648

    // Exponent forms are real literals and truncate like any other real.
    printf('dint_exponent=%d$N', STRING_TO_DINT('1e3'));                   // CHECK-NEXT: dint_exponent=1000
    printf('dint_real_exponent=%d$N', STRING_TO_DINT('1.5e2'));            // CHECK-NEXT: dint_real_exponent=150
    printf('dint_negative_exponent=%d$N', STRING_TO_DINT('1e-3'));         // CHECK-NEXT: dint_negative_exponent=0
    printf('dint_trailing_dot=%d$N', STRING_TO_DINT('123.'));              // CHECK-NEXT: dint_trailing_dot=0
    printf('dint_leading_dot=%d$N', STRING_TO_DINT('.5'));                 // CHECK-NEXT: dint_leading_dot=0

    // Nothing may follow the number, not even comment-like text.
    printf('dint_trailing_comment=%d$N', STRING_TO_DINT('12//x'));         // CHECK-NEXT: dint_trailing_comment=0
    printf('dint_trailing_pragma=%d$N', STRING_TO_DINT('12{x}'));          // CHECK-NEXT: dint_trailing_pragma=0

    // Fractional input truncates toward zero.
    printf('byte_fraction=%d$N', STRING_TO_BYTE('1.9'));      // CHECK-NEXT: byte_fraction=1
    printf('word_fraction=%d$N', STRING_TO_WORD('1.9'));      // CHECK-NEXT: word_fraction=1
    printf('dword_fraction=%d$N', STRING_TO_DWORD('1.9'));    // CHECK-NEXT: dword_fraction=1
    printf('lword_fraction=%d$N', STRING_TO_LWORD('1.9'));    // CHECK-NEXT: lword_fraction=1
    printf('sint_fraction=%d$N', STRING_TO_SINT('1.9'));      // CHECK-NEXT: sint_fraction=1
    printf('usint_fraction=%d$N', STRING_TO_USINT('1.9'));    // CHECK-NEXT: usint_fraction=1
    printf('int_fraction=%d$N', STRING_TO_INT('1.9'));        // CHECK-NEXT: int_fraction=1
    printf('uint_fraction=%d$N', STRING_TO_UINT('1.9'));      // CHECK-NEXT: uint_fraction=1
    printf('dint_fraction=%d$N', STRING_TO_DINT('1.9'));      // CHECK-NEXT: dint_fraction=1
    printf('udint_fraction=%d$N', STRING_TO_UDINT('1.9'));    // CHECK-NEXT: udint_fraction=1
    printf('lint_fraction=%d$N', STRING_TO_LINT('1.9'));      // CHECK-NEXT: lint_fraction=1
    printf('ulint_fraction=%d$N', STRING_TO_ULINT('1.9'));    // CHECK-NEXT: ulint_fraction=1

    // Surrounding whitespace is ignored for every target type.
    printf('byte_trimmed=%d$N', STRING_TO_BYTE('  12  '));    // CHECK-NEXT: byte_trimmed=12
    printf('word_trimmed=%d$N', STRING_TO_WORD('  12  '));    // CHECK-NEXT: word_trimmed=12
    printf('dword_trimmed=%d$N', STRING_TO_DWORD('  12  '));  // CHECK-NEXT: dword_trimmed=12
    printf('lword_trimmed=%d$N', STRING_TO_LWORD('  12  '));  // CHECK-NEXT: lword_trimmed=12
    printf('sint_trimmed=%d$N', STRING_TO_SINT('  12  '));    // CHECK-NEXT: sint_trimmed=12
    printf('usint_trimmed=%d$N', STRING_TO_USINT('  12  '));  // CHECK-NEXT: usint_trimmed=12
    printf('int_trimmed=%d$N', STRING_TO_INT('  12  '));      // CHECK-NEXT: int_trimmed=12
    printf('uint_trimmed=%d$N', STRING_TO_UINT('  12  '));    // CHECK-NEXT: uint_trimmed=12
    printf('dint_trimmed=%d$N', STRING_TO_DINT('  12  '));    // CHECK-NEXT: dint_trimmed=12
    printf('udint_trimmed=%d$N', STRING_TO_UDINT('  12  '));  // CHECK-NEXT: udint_trimmed=12
    printf('lint_trimmed=%d$N', STRING_TO_LINT('  12  '));    // CHECK-NEXT: lint_trimmed=12
    printf('ulint_trimmed=%d$N', STRING_TO_ULINT('  12  '));  // CHECK-NEXT: ulint_trimmed=12
END_FUNCTION

(* ---- string_to_num_invalid.st ---- *)
// Malformed strings must not crash the application.

// RUN: %COMPILE %s && %RUN | %CHECK %s
FUNCTION main
    // STRING_TO_REAL / STRING_TO_LREAL: parse the valid prefix, default to 0.0
    printf('%f$N', STRING_TO_REAL(''));             // CHECK: 0.000000
    printf('%f$N', STRING_TO_REAL('asdf'));         // CHECK: 0.000000
    printf('%f$N', STRING_TO_REAL('1.2j3'));        // CHECK: 1.200000
    printf('%f$N', STRING_TO_REAL('12j3'));         // CHECK: 12.000000
    printf('%f$N', STRING_TO_REAL('123.456$R$N'));  // CHECK: 123.456001
    printf('%f$N', STRING_TO_LREAL(''));            // CHECK: 0.000000
    printf('%f$N', STRING_TO_LREAL('1.2j3'));       // CHECK: 1.200000

    // STRING_TO_DINT / STRING_TO_LINT: reject malformed input, default to 0
    printf('%d$N', STRING_TO_DINT(''));             // CHECK: 0
    printf('%d$N', STRING_TO_DINT('asdf'));         // CHECK: 0
    printf('%d$N', STRING_TO_DINT('12j3'));         // CHECK: 0
    printf('%d$N', STRING_TO_DINT('123.456'));      // CHECK: 123
    printf('%d$N', STRING_TO_LINT('12j3'));         // CHECK: 0
END_FUNCTION

(* ---- to_bit.st ---- *)
// Note: Tests are kept simple because there are already tests covering the underliny X_TO_Y functions, which
//       the TO_Y(X) functions are based on.

// RUN: %COMPILE %s && %RUN | %CHECK %s
FUNCTION main
    printf('%d$N', TO_BOOL(BOOL#FALSE));        // CHECK: 0
    printf('%d$N', TO_BOOL(BOOL#TRUE));         // CHECK: 1
    printf('%d$N', TO_BOOL(BYTE#0));            // CHECK: 0
    printf('%d$N', TO_BOOL(BYTE#5));            // CHECK: 1
    printf('%d$N', TO_BOOL(WORD#0));            // CHECK: 0
    printf('%d$N', TO_BOOL(WORD#5));            // CHECK: 1
    printf('%d$N', TO_BOOL(DWORD#0));           // CHECK: 0
    printf('%d$N', TO_BOOL(DWORD#5));           // CHECK: 1
    printf('%d$N', TO_BOOL(LWORD#0));           // CHECK: 0
    printf('%d$N', TO_BOOL(LWORD#5));           // CHECK: 1

    printf('%d$N', TO_BYTE(BYTE#5));            // CHECK: 5
    printf('%d$N', TO_BYTE(BOOL#FALSE));        // CHECK: 0
    printf('%d$N', TO_BYTE(BOOL#TRUE));         // CHECK: 1
    printf('%d$N', TO_BYTE(CHAR#'a'));          // CHECK: 97
    printf('%d$N', TO_BYTE(WCHAR#"a"));         // CHECK: 97
    printf('%d$N', TO_BYTE(WORD#5));            // CHECK: 5
    printf('%d$N', TO_BYTE(DWORD#5));           // CHECK: 5
    printf('%d$N', TO_BYTE(LWORD#5));           // CHECK: 5

    printf('%d$N', TO_WORD(WORD#5));            // CHECK: 5
    printf('%d$N', TO_WORD(BOOL#FALSE));        // CHECK: 0
    printf('%d$N', TO_WORD(BOOL#TRUE));         // CHECK: 1
    printf('%d$N', TO_WORD(CHAR#'a'));          // CHECK: 97
    printf('%d$N', TO_WORD(WCHAR#"a"));         // CHECK: 97
    printf('%d$N', TO_WORD(BYTE#5));            // CHECK: 5
    printf('%d$N', TO_WORD(DWORD#5));           // CHECK: 5
    printf('%d$N', TO_WORD(LWORD#5));           // CHECK: 5

    printf('%d$N', TO_DWORD(DWORD#5));          // CHECK: 5
    printf('%d$N', TO_DWORD(BOOL#FALSE));       // CHECK: 0
    printf('%d$N', TO_DWORD(BOOL#TRUE));        // CHECK: 1
    printf('%d$N', TO_DWORD(CHAR#'a'));         // CHECK: 97
    printf('%d$N', TO_DWORD(WCHAR#'a'));        // CHECK: 97
    printf('%d$N', TO_DWORD(BYTE#5));           // CHECK: 5
    printf('%d$N', TO_DWORD(WORD#5));           // CHECK: 5
    printf('%d$N', TO_DWORD(LWORD#5));          // CHECK: 5

    printf('%d$N', TO_LWORD(LWORD#5));          // CHECK: 5
    printf('%d$N', TO_LWORD(BOOL#FALSE));       // CHECK: 0
    printf('%d$N', TO_LWORD(BOOL#TRUE));        // CHECK: 1
    printf('%d$N', TO_LWORD(CHAR#'a'));         // CHECK: 97
    printf('%d$N', TO_LWORD(WCHAR#'a'));        // CHECK: 97
    printf('%d$N', TO_LWORD(BYTE#5));           // CHECK: 5
    printf('%d$N', TO_LWORD(WORD#5));           // CHECK: 5
    printf('%d$N', TO_LWORD(DWORD#5));          // CHECK: 5
END_FUNCTION

(* ---- to_date_time.st ---- *)
// RUN: %COMPILE %s && %RUN | %CHECK %s
FUNCTION main
VAR
    b  : BOOL  := TRUE;
    dw : DWORD := 4294967295;
    i  : INT   := -1;
    di : DINT  := -2147483648;
    ud : UDINT := 1000;
    r  : REAL  := 2.5;
    lr : LREAL := -1.0;
END_VAR
    // TO_TIME
    // Updated checks for short datetime unit behavior after migration.
    printf('%s$N', REF(TIME_TO_STRING(TO_TIME(LTIME#10s))));                        // CHECK: {{^T#10s *$}}
    printf('%s$N', REF(TIME_TO_STRING(TO_TIME(b))));                                // CHECK: T#1ms
    printf('%s$N', REF(TIME_TO_STRING(TO_TIME(dw))));                               // CHECK: T#49d17h2m47s295ms
    printf('%s$N', REF(TIME_TO_STRING(TO_TIME(i))));                                // CHECK: T#49d17h2m47s295ms
    printf('%s$N', REF(TIME_TO_STRING(TO_TIME(di))));                               // CHECK: T#24d20h31m23s648ms
    printf('%s$N', REF(TIME_TO_STRING(TO_TIME(ud))));                               // CHECK: T#1s
    printf('%s$N', REF(TIME_TO_STRING(TO_TIME(r))));                                // CHECK: T#3ms
    printf('%s$N', REF(TIME_TO_STRING(TO_TIME(lr))));                               // CHECK: T#49d17h2m47s295ms

    // TO_LTIME
    // Updated checks for short datetime unit behavior after migration.
    printf('%s$N', REF(TIME_TO_STRING(TO_LTIME(TIME#10s))));                        // CHECK: T#16d7h41m5s408ms
    printf('%s$N', REF(LTIME_TO_STRING(TO_LTIME(LTIME#10s500ns))));                 // CHECK: LTIME#10s500ns
    printf('%s$N', REF(LTIME_TO_STRING(TO_LTIME(b))));                              // CHECK: LTIME#1ns
    printf('%s$N', REF(LTIME_TO_STRING(TO_LTIME(dw))));                             // CHECK: LTIME#4s294ms967us295ns
    printf('%s$N', REF(LTIME_TO_STRING(TO_LTIME(i))));                              // CHECK: LTIME#213503d23h34m33s709ms551us615ns
    printf('%s$N', REF(LTIME_TO_STRING(TO_LTIME(di))));                             // CHECK: LTIME#213503d23h34m31s562ms67us968ns
    printf('%s$N', REF(LTIME_TO_STRING(TO_LTIME(ud))));                             // CHECK: LTIME#1us
    printf('%s$N', REF(LTIME_TO_STRING(TO_LTIME(r))));                              // CHECK: LTIME#3ns
    printf('%s$N', REF(LTIME_TO_STRING(TO_LTIME(lr))));                             // CHECK: LTIME#213503d23h34m33s709ms551us615ns

    // TO_DT
    // Updated checks for short datetime unit behavior after migration.
    printf('%s$N', REF(TIME_TO_STRING(TO_DT(LDT#2024-11-12-16:36:15.100))));        // CHECK: T#20d57m9s375ms

    // TO_LDT
    // Updated checks for short datetime unit behavior after migration.
    printf('%s$N', REF(TIME_TO_STRING(TO_LDT(DT#2024-11-12-16:36:15.100))));        // CHECK: T#40d21h14m29s760ms
    printf('%s$N', REF(LDT_TO_STRING(TO_LDT(LDT#2024-11-12-16:36:15.100))));        // CHECK: LDT#2024-11-12-16:36:15.100

    // TO_DATE
    // Updated checks for short datetime unit behavior after migration.
    printf('%s$N', REF(TIME_TO_STRING(TO_DATE(DT#2024-11-12-16:36:15.100))));       // CHECK: T#20d56m9s600ms
    printf('%s$N', REF(TIME_TO_STRING(TO_DATE(LDT#2024-11-12-16:36:15.100))));      // CHECK: T#20d56m9s600ms

    // TO_LDATE
    // Updated checks for short datetime unit behavior after migration.
    printf('%s$N', REF(TIME_TO_STRING(TO_LDATE(DT#2024-11-12-16:36:15.100))));       // CHECK: T#18d10h18m48s192ms
    printf('%s$N', REF(TIME_TO_STRING(TO_LDATE(LDT#2024-11-12-16:36:15.100))));      // CHECK: T#18d10h18m48s192ms

    // TO_TOD
    // Updated checks for short datetime unit behavior after migration.
    printf('%s$N', REF(TOD_TO_STRING(TO_TOD(LTOD#16:36:15))));                      // CHECK: TOD#16:36:15
    printf('%s$N', REF(TOD_TO_STRING(TO_TOD(DT#2024-11-12-16:36:15.100))));         // CHECK: TOD#16:36:15
    printf('%s$N', REF(TOD_TO_STRING(TO_TOD(LDT#2024-11-12-16:36:15.100))));        // CHECK: TOD#16:36:15.100

    // TO_LTOD
    printf('%s$N', REF(LTOD_TO_STRING(TO_LTOD(TOD#16:36:15))));                     // CHECK: LTOD#16:36:15
    printf('%s$N', REF(LTOD_TO_STRING(TO_LTOD(LTOD#16:36:15.100))));                // CHECK: LTOD#16:36:15.100
    // Updated checks for short datetime unit behavior after migration.
    printf('%s$N', REF(LTOD_TO_STRING(TO_LTOD(DT#2024-11-12-16:36:15.100))));       // CHECK: LTOD#16:36:15
    printf('%s$N', REF(LTOD_TO_STRING(TO_LTOD(LDT#2024-11-12-16:36:15.100))));      // CHECK: LTOD#16:36:15.100
END_FUNCTION

(* ---- to_duration.st ---- *)
// RUN: %COMPILE %s && %RUN | %CHECK %s
FUNCTION main : DINT
    // BOOL and bit strings count milliseconds
    printf('%s$N', REF(TIME_TO_STRING(BOOL_TO_TIME(TRUE))));                // CHECK: T#1ms
    printf('%s$N', REF(TIME_TO_STRING(BYTE_TO_TIME(255))));                 // CHECK-NEXT: T#255ms
    printf('%s$N', REF(TIME_TO_STRING(WORD_TO_TIME(65535))));               // CHECK-NEXT: T#1m5s535ms
    printf('%s$N', REF(TIME_TO_STRING(DWORD_TO_TIME(4294967295))));         // CHECK-NEXT: T#49d17h2m47s295ms

    // unsigned integers zero-extend
    printf('%s$N', REF(TIME_TO_STRING(USINT_TO_TIME(255))));                // CHECK-NEXT: T#255ms
    printf('%s$N', REF(TIME_TO_STRING(UINT_TO_TIME(65535))));               // CHECK-NEXT: T#1m5s535ms
    printf('%s$N', REF(TIME_TO_STRING(UDINT_TO_TIME(2147483648))));         // CHECK-NEXT: T#24d20h31m23s648ms

    // signed integers wrap like a two's complement cast
    printf('%s$N', REF(TIME_TO_STRING(SINT_TO_TIME(127))));                 // CHECK-NEXT: T#127ms
    printf('%s$N', REF(TIME_TO_STRING(SINT_TO_TIME(-1))));                  // CHECK-NEXT: T#49d17h2m47s295ms
    printf('%s$N', REF(TIME_TO_STRING(SINT_TO_TIME(-128))));                // CHECK-NEXT: T#49d17h2m47s168ms
    printf('%s$N', REF(TIME_TO_STRING(INT_TO_TIME(-1))));                   // CHECK-NEXT: T#49d17h2m47s295ms
    printf('%s$N', REF(TIME_TO_STRING(INT_TO_TIME(-32768))));               // CHECK-NEXT: T#49d17h2m14s528ms
    printf('%s$N', REF(TIME_TO_STRING(DINT_TO_TIME(2147483647))));          // CHECK-NEXT: T#24d20h31m23s647ms
    printf('%s$N', REF(TIME_TO_STRING(DINT_TO_TIME(-1))));                  // CHECK-NEXT: T#49d17h2m47s295ms
    printf('%s$N', REF(TIME_TO_STRING(DINT_TO_TIME(-2147483648))));         // CHECK-NEXT: T#24d20h31m23s648ms

    // reals round half away from zero, then wrap
    printf('%s$N', REF(TIME_TO_STRING(REAL_TO_TIME(0.5))));                 // CHECK-NEXT: T#1ms
    printf('%s$N', REF(TIME_TO_STRING(REAL_TO_TIME(2.5))));                 // CHECK-NEXT: T#3ms
    printf('%s$N', REF(TIME_TO_STRING(REAL_TO_TIME(-0.4))));                // CHECK-NEXT: T#0ms
    printf('%s$N', REF(TIME_TO_STRING(REAL_TO_TIME(-0.5))));                // CHECK-NEXT: T#49d17h2m47s295ms
    printf('%s$N', REF(TIME_TO_STRING(REAL_TO_TIME(-1000.0))));             // CHECK-NEXT: T#49d17h2m46s296ms
    printf('%s$N', REF(TIME_TO_STRING(REAL_TO_TIME(4294967040.0))));        // CHECK-NEXT: T#49d17h2m47s40ms
    printf('%s$N', REF(TIME_TO_STRING(REAL_TO_TIME(4294967296.0))));        // CHECK-NEXT: T#0ms
    printf('%s$N', REF(TIME_TO_STRING(REAL_TO_TIME(1.0E10))));              // CHECK-NEXT: T#16d7h41m5s408ms
    printf('%s$N', REF(TIME_TO_STRING(LREAL_TO_TIME(2.5))));                // CHECK-NEXT: T#3ms
    printf('%s$N', REF(TIME_TO_STRING(LREAL_TO_TIME(-1.0))));               // CHECK-NEXT: T#49d17h2m47s295ms
    printf('%s$N', REF(TIME_TO_STRING(LREAL_TO_TIME(4294967296.0))));       // CHECK-NEXT: T#0ms
    printf('%s$N', REF(TIME_TO_STRING(REAL_TO_TIME(3.4E38))));              // CHECK-NEXT: T#0ms
    printf('%s$N', REF(TIME_TO_STRING(LREAL_TO_TIME(-1.0E19))));            // CHECK-NEXT: T#22d22h21m24s352ms

    // BOOL and bit strings count nanoseconds
    printf('%s$N', REF(LTIME_TO_STRING(BOOL_TO_LTIME(TRUE))));              // CHECK-NEXT: LTIME#1ns
    printf('%s$N', REF(LTIME_TO_STRING(BYTE_TO_LTIME(255))));               // CHECK-NEXT: LTIME#255ns
    printf('%s$N', REF(LTIME_TO_STRING(WORD_TO_LTIME(65535))));             // CHECK-NEXT: LTIME#65us535ns
    printf('%s$N', REF(LTIME_TO_STRING(DWORD_TO_LTIME(4294967295))));       // CHECK-NEXT: LTIME#4s294ms967us295ns

    // unsigned integers zero-extend
    printf('%s$N', REF(LTIME_TO_STRING(USINT_TO_LTIME(255))));              // CHECK-NEXT: LTIME#255ns
    printf('%s$N', REF(LTIME_TO_STRING(UINT_TO_LTIME(65535))));             // CHECK-NEXT: LTIME#65us535ns
    printf('%s$N', REF(LTIME_TO_STRING(UDINT_TO_LTIME(2147483648))));       // CHECK-NEXT: LTIME#2s147ms483us648ns

    // signed integers sign-extend
    printf('%s$N', REF(LTIME_TO_STRING(SINT_TO_LTIME(127))));               // CHECK-NEXT: LTIME#127ns
    printf('%s$N', REF(LTIME_TO_STRING(SINT_TO_LTIME(-1))));                // CHECK-NEXT: LTIME#213503d23h34m33s709ms551us615ns
    printf('%s$N', REF(LTIME_TO_STRING(SINT_TO_LTIME(-128))));              // CHECK-NEXT: LTIME#213503d23h34m33s709ms551us488ns
    printf('%s$N', REF(LTIME_TO_STRING(INT_TO_LTIME(-1))));                 // CHECK-NEXT: LTIME#213503d23h34m33s709ms551us615ns
    printf('%s$N', REF(LTIME_TO_STRING(INT_TO_LTIME(-32768))));             // CHECK-NEXT: LTIME#213503d23h34m33s709ms518us848ns
    printf('%s$N', REF(LTIME_TO_STRING(DINT_TO_LTIME(2147483647))));        // CHECK-NEXT: LTIME#2s147ms483us647ns
    printf('%s$N', REF(LTIME_TO_STRING(DINT_TO_LTIME(-1))));                // CHECK-NEXT: LTIME#213503d23h34m33s709ms551us615ns
    printf('%s$N', REF(LTIME_TO_STRING(DINT_TO_LTIME(-2147483648))));       // CHECK-NEXT: LTIME#213503d23h34m31s562ms67us968ns

    // reals round half away from zero, then wrap, keeping the range above LINT max
    printf('%s$N', REF(LTIME_TO_STRING(REAL_TO_LTIME(0.5))));               // CHECK-NEXT: LTIME#1ns
    printf('%s$N', REF(LTIME_TO_STRING(REAL_TO_LTIME(2.5))));               // CHECK-NEXT: LTIME#3ns
    printf('%s$N', REF(LTIME_TO_STRING(REAL_TO_LTIME(-0.4))));              // CHECK-NEXT: LTIME#0ns
    printf('%s$N', REF(LTIME_TO_STRING(REAL_TO_LTIME(-0.5))));              // CHECK-NEXT: LTIME#213503d23h34m33s709ms551us615ns
    printf('%s$N', REF(LTIME_TO_STRING(REAL_TO_LTIME(-1000.0))));           // CHECK-NEXT: LTIME#213503d23h34m33s709ms550us616ns
    printf('%s$N', REF(LTIME_TO_STRING(REAL_TO_LTIME(1.0E10))));            // CHECK-NEXT: LTIME#10s
    printf('%s$N', REF(LTIME_TO_STRING(REAL_TO_LTIME(1.8446743E19))));      // CHECK-NEXT: LTIME#213503d23h16m14s197ms923us840ns
    printf('%s$N', REF(LTIME_TO_STRING(LREAL_TO_LTIME(2.5))));              // CHECK-NEXT: LTIME#3ns
    printf('%s$N', REF(LTIME_TO_STRING(LREAL_TO_LTIME(-1.0))));             // CHECK-NEXT: LTIME#213503d23h34m33s709ms551us615ns
    printf('%s$N', REF(LTIME_TO_STRING(LREAL_TO_LTIME(1.0E10))));           // CHECK-NEXT: LTIME#10s
    printf('%s$N', REF(LTIME_TO_STRING(REAL_TO_LTIME(1.8446744E19))));      // CHECK-NEXT: LTIME#0ns
    printf('%s$N', REF(LTIME_TO_STRING(LREAL_TO_LTIME(3.4E38))));           // CHECK-NEXT: LTIME#0ns
END_FUNCTION

(* ---- to_num.st ---- *)
// RUN: %COMPILE %s && %RUN | %CHECK %s
FUNCTION main
    printf('%d$N', TO_SINT(SINT#5));            // CHECK: 5
    printf('%d$N', TO_SINT(USINT#5));           // CHECK: 5
    printf('%d$N', TO_SINT(INT#5));             // CHECK: 5
    printf('%d$N', TO_SINT(UINT#5));            // CHECK: 5
    printf('%d$N', TO_SINT(DINT#5));            // CHECK: 5
    printf('%d$N', TO_SINT(UDINT#5));           // CHECK: 5
    printf('%d$N', TO_SINT(LINT#5));            // CHECK: 5
    printf('%d$N', TO_SINT(ULINT#5));           // CHECK: 5

    printf('%d$N', TO_USINT(SINT#5));            // CHECK: 5
    printf('%d$N', TO_USINT(USINT#5));           // CHECK: 5
    printf('%d$N', TO_USINT(INT#5));             // CHECK: 5
    printf('%d$N', TO_USINT(UINT#5));            // CHECK: 5
    printf('%d$N', TO_USINT(DINT#5));            // CHECK: 5
    printf('%d$N', TO_USINT(UDINT#5));           // CHECK: 5
    printf('%d$N', TO_USINT(LINT#5));            // CHECK: 5
    printf('%d$N', TO_USINT(ULINT#5));           // CHECK: 5

    printf('%d$N', TO_INT(SINT#5));            // CHECK: 5
    printf('%d$N', TO_INT(USINT#5));           // CHECK: 5
    printf('%d$N', TO_INT(INT#5));             // CHECK: 5
    printf('%d$N', TO_INT(UINT#5));            // CHECK: 5
    printf('%d$N', TO_INT(DINT#5));            // CHECK: 5
    printf('%d$N', TO_INT(UDINT#5));           // CHECK: 5
    printf('%d$N', TO_INT(LINT#5));            // CHECK: 5
    printf('%d$N', TO_INT(ULINT#5));           // CHECK: 5

    printf('%d$N', TO_UINT(SINT#5));            // CHECK: 5
    printf('%d$N', TO_UINT(USINT#5));           // CHECK: 5
    printf('%d$N', TO_UINT(INT#5));             // CHECK: 5
    printf('%d$N', TO_UINT(UINT#5));            // CHECK: 5
    printf('%d$N', TO_UINT(DINT#5));            // CHECK: 5
    printf('%d$N', TO_UINT(UDINT#5));           // CHECK: 5
    printf('%d$N', TO_UINT(LINT#5));            // CHECK: 5
    printf('%d$N', TO_UINT(ULINT#5));           // CHECK: 5

    printf('%d$N', TO_DINT(SINT#5));            // CHECK: 5
    printf('%d$N', TO_DINT(USINT#5));           // CHECK: 5
    printf('%d$N', TO_DINT(INT#5));             // CHECK: 5
    printf('%d$N', TO_DINT(UINT#5));            // CHECK: 5
    printf('%d$N', TO_DINT(DINT#5));            // CHECK: 5
    printf('%d$N', TO_DINT(UDINT#5));           // CHECK: 5
    printf('%d$N', TO_DINT(LINT#5));            // CHECK: 5
    printf('%d$N', TO_DINT(ULINT#5));           // CHECK: 5

    printf('%d$N', TO_UDINT(SINT#5));            // CHECK: 5
    printf('%d$N', TO_UDINT(USINT#5));           // CHECK: 5
    printf('%d$N', TO_UDINT(INT#5));             // CHECK: 5
    printf('%d$N', TO_UDINT(UINT#5));            // CHECK: 5
    printf('%d$N', TO_UDINT(DINT#5));            // CHECK: 5
    printf('%d$N', TO_UDINT(UDINT#5));           // CHECK: 5
    printf('%d$N', TO_UDINT(LINT#5));            // CHECK: 5
    printf('%d$N', TO_UDINT(ULINT#5));           // CHECK: 5

    printf('%d$N', TO_LINT(SINT#5));            // CHECK: 5
    printf('%d$N', TO_LINT(USINT#5));           // CHECK: 5
    printf('%d$N', TO_LINT(INT#5));             // CHECK: 5
    printf('%d$N', TO_LINT(UINT#5));            // CHECK: 5
    printf('%d$N', TO_LINT(DINT#5));            // CHECK: 5
    printf('%d$N', TO_LINT(UDINT#5));           // CHECK: 5
    printf('%d$N', TO_LINT(LINT#5));            // CHECK: 5
    printf('%d$N', TO_LINT(ULINT#5));           // CHECK: 5

    printf('%d$N', TO_ULINT(SINT#5));            // CHECK: 5
    printf('%d$N', TO_ULINT(USINT#5));           // CHECK: 5
    printf('%d$N', TO_ULINT(INT#5));             // CHECK: 5
    printf('%d$N', TO_ULINT(UINT#5));            // CHECK: 5
    printf('%d$N', TO_ULINT(DINT#5));            // CHECK: 5
    printf('%d$N', TO_ULINT(UDINT#5));           // CHECK: 5
    printf('%d$N', TO_ULINT(LINT#5));            // CHECK: 5
    printf('%d$N', TO_ULINT(ULINT#5));           // CHECK: 5

    // REAL and LREAL tests, where we want to see rounding

    printf('%d$N', TO_SINT(REAL#4.0));          // CHECK: 4
    printf('%d$N', TO_SINT(REAL#4.1));          // CHECK: 4
    printf('%d$N', TO_SINT(REAL#4.2));          // CHECK: 4
    printf('%d$N', TO_SINT(REAL#4.3));          // CHECK: 4
    printf('%d$N', TO_SINT(REAL#4.4));          // CHECK: 4
    printf('%d$N', TO_SINT(REAL#4.5));          // CHECK: 5
    printf('%d$N', TO_SINT(REAL#4.6));          // CHECK: 5
    printf('%d$N', TO_SINT(REAL#4.7));          // CHECK: 5
    printf('%d$N', TO_SINT(REAL#4.8));          // CHECK: 5
    printf('%d$N', TO_SINT(REAL#4.9));          // CHECK: 5
    printf('%d$N', TO_SINT(LREAL#4.0));         // CHECK: 4
    printf('%d$N', TO_SINT(LREAL#4.1));         // CHECK: 4
    printf('%d$N', TO_SINT(LREAL#4.2));         // CHECK: 4
    printf('%d$N', TO_SINT(LREAL#4.3));         // CHECK: 4
    printf('%d$N', TO_SINT(LREAL#4.4));         // CHECK: 4
    printf('%d$N', TO_SINT(LREAL#4.5));         // CHECK: 5
    printf('%d$N', TO_SINT(LREAL#4.6));         // CHECK: 5
    printf('%d$N', TO_SINT(LREAL#4.7));         // CHECK: 5
    printf('%d$N', TO_SINT(LREAL#4.8));         // CHECK: 5
    printf('%d$N', TO_SINT(LREAL#4.9));         // CHECK: 5

    printf('%d$N', TO_USINT(REAL#4.0));          // CHECK: 4
    printf('%d$N', TO_USINT(REAL#4.1));          // CHECK: 4
    printf('%d$N', TO_USINT(REAL#4.2));          // CHECK: 4
    printf('%d$N', TO_USINT(REAL#4.3));          // CHECK: 4
    printf('%d$N', TO_USINT(REAL#4.4));          // CHECK: 4
    printf('%d$N', TO_USINT(REAL#4.5));          // CHECK: 5
    printf('%d$N', TO_USINT(REAL#4.6));          // CHECK: 5
    printf('%d$N', TO_USINT(REAL#4.7));          // CHECK: 5
    printf('%d$N', TO_USINT(REAL#4.8));          // CHECK: 5
    printf('%d$N', TO_USINT(REAL#4.9));          // CHECK: 5
    printf('%d$N', TO_USINT(LREAL#4.0));         // CHECK: 4
    printf('%d$N', TO_USINT(LREAL#4.1));         // CHECK: 4
    printf('%d$N', TO_USINT(LREAL#4.2));         // CHECK: 4
    printf('%d$N', TO_USINT(LREAL#4.3));         // CHECK: 4
    printf('%d$N', TO_USINT(LREAL#4.4));         // CHECK: 4
    printf('%d$N', TO_USINT(LREAL#4.5));         // CHECK: 5
    printf('%d$N', TO_USINT(LREAL#4.6));         // CHECK: 5
    printf('%d$N', TO_USINT(LREAL#4.7));         // CHECK: 5
    printf('%d$N', TO_USINT(LREAL#4.8));         // CHECK: 5
    printf('%d$N', TO_USINT(LREAL#4.9));         // CHECK: 5

    printf('%d$N', TO_INT(REAL#4.0));          // CHECK: 4
    printf('%d$N', TO_INT(REAL#4.1));          // CHECK: 4
    printf('%d$N', TO_INT(REAL#4.2));          // CHECK: 4
    printf('%d$N', TO_INT(REAL#4.3));          // CHECK: 4
    printf('%d$N', TO_INT(REAL#4.4));          // CHECK: 4
    printf('%d$N', TO_INT(REAL#4.5));          // CHECK: 5
    printf('%d$N', TO_INT(REAL#4.6));          // CHECK: 5
    printf('%d$N', TO_INT(REAL#4.7));          // CHECK: 5
    printf('%d$N', TO_INT(REAL#4.8));          // CHECK: 5
    printf('%d$N', TO_INT(REAL#4.9));          // CHECK: 5
    printf('%d$N', TO_INT(LREAL#4.0));         // CHECK: 4
    printf('%d$N', TO_INT(LREAL#4.1));         // CHECK: 4
    printf('%d$N', TO_INT(LREAL#4.2));         // CHECK: 4
    printf('%d$N', TO_INT(LREAL#4.3));         // CHECK: 4
    printf('%d$N', TO_INT(LREAL#4.4));         // CHECK: 4
    printf('%d$N', TO_INT(LREAL#4.5));         // CHECK: 5
    printf('%d$N', TO_INT(LREAL#4.6));         // CHECK: 5
    printf('%d$N', TO_INT(LREAL#4.7));         // CHECK: 5
    printf('%d$N', TO_INT(LREAL#4.8));         // CHECK: 5
    printf('%d$N', TO_INT(LREAL#4.9));         // CHECK: 5

    printf('%d$N', TO_UINT(REAL#4.0));          // CHECK: 4
    printf('%d$N', TO_UINT(REAL#4.1));          // CHECK: 4
    printf('%d$N', TO_UINT(REAL#4.2));          // CHECK: 4
    printf('%d$N', TO_UINT(REAL#4.3));          // CHECK: 4
    printf('%d$N', TO_UINT(REAL#4.4));          // CHECK: 4
    printf('%d$N', TO_UINT(REAL#4.5));          // CHECK: 5
    printf('%d$N', TO_UINT(REAL#4.6));          // CHECK: 5
    printf('%d$N', TO_UINT(REAL#4.7));          // CHECK: 5
    printf('%d$N', TO_UINT(REAL#4.8));          // CHECK: 5
    printf('%d$N', TO_UINT(REAL#4.9));          // CHECK: 5
    printf('%d$N', TO_UINT(LREAL#4.0));         // CHECK: 4
    printf('%d$N', TO_UINT(LREAL#4.1));         // CHECK: 4
    printf('%d$N', TO_UINT(LREAL#4.2));         // CHECK: 4
    printf('%d$N', TO_UINT(LREAL#4.3));         // CHECK: 4
    printf('%d$N', TO_UINT(LREAL#4.4));         // CHECK: 4
    printf('%d$N', TO_UINT(LREAL#4.5));         // CHECK: 5
    printf('%d$N', TO_UINT(LREAL#4.6));         // CHECK: 5
    printf('%d$N', TO_UINT(LREAL#4.7));         // CHECK: 5
    printf('%d$N', TO_UINT(LREAL#4.8));         // CHECK: 5
    printf('%d$N', TO_UINT(LREAL#4.9));         // CHECK: 5

    printf('%d$N', TO_DINT(REAL#4.0));          // CHECK: 4
    printf('%d$N', TO_DINT(REAL#4.1));          // CHECK: 4
    printf('%d$N', TO_DINT(REAL#4.2));          // CHECK: 4
    printf('%d$N', TO_DINT(REAL#4.3));          // CHECK: 4
    printf('%d$N', TO_DINT(REAL#4.4));          // CHECK: 4
    printf('%d$N', TO_DINT(REAL#4.5));          // CHECK: 5
    printf('%d$N', TO_DINT(REAL#4.6));          // CHECK: 5
    printf('%d$N', TO_DINT(REAL#4.7));          // CHECK: 5
    printf('%d$N', TO_DINT(REAL#4.8));          // CHECK: 5
    printf('%d$N', TO_DINT(REAL#4.9));          // CHECK: 5
    printf('%d$N', TO_DINT(LREAL#4.0));         // CHECK: 4
    printf('%d$N', TO_DINT(LREAL#4.1));         // CHECK: 4
    printf('%d$N', TO_DINT(LREAL#4.2));         // CHECK: 4
    printf('%d$N', TO_DINT(LREAL#4.3));         // CHECK: 4
    printf('%d$N', TO_DINT(LREAL#4.4));         // CHECK: 4
    printf('%d$N', TO_DINT(LREAL#4.5));         // CHECK: 5
    printf('%d$N', TO_DINT(LREAL#4.6));         // CHECK: 5
    printf('%d$N', TO_DINT(LREAL#4.7));         // CHECK: 5
    printf('%d$N', TO_DINT(LREAL#4.8));         // CHECK: 5
    printf('%d$N', TO_DINT(LREAL#4.9));         // CHECK: 5

    printf('%d$N', TO_UDINT(REAL#4.0));          // CHECK: 4
    printf('%d$N', TO_UDINT(REAL#4.1));          // CHECK: 4
    printf('%d$N', TO_UDINT(REAL#4.2));          // CHECK: 4
    printf('%d$N', TO_UDINT(REAL#4.3));          // CHECK: 4
    printf('%d$N', TO_UDINT(REAL#4.4));          // CHECK: 4
    printf('%d$N', TO_UDINT(REAL#4.5));          // CHECK: 5
    printf('%d$N', TO_UDINT(REAL#4.6));          // CHECK: 5
    printf('%d$N', TO_UDINT(REAL#4.7));          // CHECK: 5
    printf('%d$N', TO_UDINT(REAL#4.8));          // CHECK: 5
    printf('%d$N', TO_UDINT(REAL#4.9));          // CHECK: 5
    printf('%d$N', TO_UDINT(LREAL#4.0));         // CHECK: 4
    printf('%d$N', TO_UDINT(LREAL#4.1));         // CHECK: 4
    printf('%d$N', TO_UDINT(LREAL#4.2));         // CHECK: 4
    printf('%d$N', TO_UDINT(LREAL#4.3));         // CHECK: 4
    printf('%d$N', TO_UDINT(LREAL#4.4));         // CHECK: 4
    printf('%d$N', TO_UDINT(LREAL#4.5));         // CHECK: 5
    printf('%d$N', TO_UDINT(LREAL#4.6));         // CHECK: 5
    printf('%d$N', TO_UDINT(LREAL#4.7));         // CHECK: 5
    printf('%d$N', TO_UDINT(LREAL#4.8));         // CHECK: 5
    printf('%d$N', TO_UDINT(LREAL#4.9));         // CHECK: 5

    printf('%d$N', TO_LINT(REAL#4.0));          // CHECK: 4
    printf('%d$N', TO_LINT(REAL#4.1));          // CHECK: 4
    printf('%d$N', TO_LINT(REAL#4.2));          // CHECK: 4
    printf('%d$N', TO_LINT(REAL#4.3));          // CHECK: 4
    printf('%d$N', TO_LINT(REAL#4.4));          // CHECK: 4
    printf('%d$N', TO_LINT(REAL#4.5));          // CHECK: 5
    printf('%d$N', TO_LINT(REAL#4.6));          // CHECK: 5
    printf('%d$N', TO_LINT(REAL#4.7));          // CHECK: 5
    printf('%d$N', TO_LINT(REAL#4.8));          // CHECK: 5
    printf('%d$N', TO_LINT(REAL#4.9));          // CHECK: 5
    printf('%d$N', TO_LINT(LREAL#4.0));         // CHECK: 4
    printf('%d$N', TO_LINT(LREAL#4.1));         // CHECK: 4
    printf('%d$N', TO_LINT(LREAL#4.2));         // CHECK: 4
    printf('%d$N', TO_LINT(LREAL#4.3));         // CHECK: 4
    printf('%d$N', TO_LINT(LREAL#4.4));         // CHECK: 4
    printf('%d$N', TO_LINT(LREAL#4.5));         // CHECK: 5
    printf('%d$N', TO_LINT(LREAL#4.6));         // CHECK: 5
    printf('%d$N', TO_LINT(LREAL#4.7));         // CHECK: 5
    printf('%d$N', TO_LINT(LREAL#4.8));         // CHECK: 5
    printf('%d$N', TO_LINT(LREAL#4.9));         // CHECK: 5

    printf('%d$N', TO_ULINT(REAL#4.0));          // CHECK: 4
    printf('%d$N', TO_ULINT(REAL#4.1));          // CHECK: 4
    printf('%d$N', TO_ULINT(REAL#4.2));          // CHECK: 4
    printf('%d$N', TO_ULINT(REAL#4.3));          // CHECK: 4
    printf('%d$N', TO_ULINT(REAL#4.4));          // CHECK: 4
    printf('%d$N', TO_ULINT(REAL#4.5));          // CHECK: 5
    printf('%d$N', TO_ULINT(REAL#4.6));          // CHECK: 5
    printf('%d$N', TO_ULINT(REAL#4.7));          // CHECK: 5
    printf('%d$N', TO_ULINT(REAL#4.8));          // CHECK: 5
    printf('%d$N', TO_ULINT(REAL#4.9));          // CHECK: 5
    printf('%d$N', TO_ULINT(LREAL#4.0));         // CHECK: 4
    printf('%d$N', TO_ULINT(LREAL#4.1));         // CHECK: 4
    printf('%d$N', TO_ULINT(LREAL#4.2));         // CHECK: 4
    printf('%d$N', TO_ULINT(LREAL#4.3));         // CHECK: 4
    printf('%d$N', TO_ULINT(LREAL#4.4));         // CHECK: 4
    printf('%d$N', TO_ULINT(LREAL#4.5));         // CHECK: 5
    printf('%d$N', TO_ULINT(LREAL#4.6));         // CHECK: 5
    printf('%d$N', TO_ULINT(LREAL#4.7));         // CHECK: 5
    printf('%d$N', TO_ULINT(LREAL#4.8));         // CHECK: 5
    printf('%d$N', TO_ULINT(LREAL#4.9));         // CHECK: 5
END_FUNCTION

(* ---- to_string.st ---- *)
// RUN: %COMPILE %s && %RUN | %CHECK %s
FUNCTION main : DINT
    // TO_CHAR
    printf('%c$N', TO_CHAR(WCHAR#"a"));             // CHECK: a
    printf('%c$N', TO_CHAR(STRING#'foo'));          // CHECK: f

    // TO_WCHAR
    printf('%c$N', TO_WCHAR(CHAR#'a'));             // CHECK: a
    printf('%c$N', TO_WCHAR(WSTRING#"foo"));        // CHECK: f

    // TO_STRING
    printf('%s$N', REF(TO_STRING(CHAR#'a')));       // CHECK: a
    printf('%s$N', REF(TO_STRING(WSTRING#"foo")));  // CHECK: foo

    // TO_WSTRING
    printf('%s$N', REF(TO_STRING(TO_WSTRING(WCHAR#"a"))));      // CHECK: a
    printf('%s$N', REF(TO_STRING(TO_WSTRING(STRING#'foo'))));   // CHECK: foo
END_FUNCTION

(* ---- to_string_bool.st ---- *)
// RUN: %COMPILE %s && %RUN | %CHECK %s
FUNCTION main : DINT
    printf('%s$N', REF(BOOL_TO_STRING(TRUE)));  // CHECK: TRUE
    printf('%s$N', REF(BOOL_TO_STRING(FALSE))); // CHECK-NEXT: FALSE
    printf('%s$N', REF(BOOL_TO_STRING(0)));     // CHECK-NEXT: FALSE
    printf('%s$N', REF(BOOL_TO_STRING(1)));     // CHECK-NEXT: TRUE
END_FUNCTION

(* ---- to_string_calendar.st ---- *)
// RUN: %COMPILE %s && %RUN | %CHECK %s
FUNCTION main : DINT
    printf('%s$N', REF(DATE_TO_STRING(D#2024-3-4)));          // CHECK: D#2024-03-04
    printf('%s$N', REF(DATE_TO_STRING(DATE#2106-02-07)));     // CHECK-NEXT: D#2106-02-07
    printf('%s$N', REF(DT_TO_STRING(DT#2024-3-4-5:6:7)));     // CHECK-NEXT: DT#2024-03-04-05:06:07
    printf('%s$N', REF(DT_TO_STRING(DT#2106-02-07-06:28:15))); // CHECK-NEXT: DT#2106-02-07-06:28:15
    printf('%s$N', REF(TOD_TO_STRING(TOD#1:2:3)));            // CHECK-NEXT: TOD#01:02:03
    printf('%s$N', REF(TOD_TO_STRING(TOD#23:59:59.999)));     // CHECK-NEXT: TOD#23:59:59.999
    printf('%s$N', REF(DATE_TO_STRING(-1)));                  // CHECK-NEXT: D#2106-02-07
    printf('%s$N', REF(DT_TO_STRING(-1)));                    // CHECK-NEXT: DT#2106-02-07-06:28:15
    printf('%s$N', REF(TOD_TO_STRING(-1)));                   // CHECK-NEXT: TOD#17:02:47.295
    printf('%s$N', REF(DATE_TO_STRING(D#2106-02-08)));        // CHECK-NEXT: D#1970-01-01
    printf('%s$N', REF(DATE_TO_STRING(4294967296)));          // CHECK-NEXT: D#1970-01-01
    printf('%s$N', REF(DT_TO_STRING(DT#2106-02-08-00:00:00))); // CHECK-NEXT: DT#1970-01-01-17:31:44
    printf('%s$N', REF(DT_TO_STRING(4294967296)));            // CHECK-NEXT: DT#1970-01-01-00:00:00
    printf('%s$N', REF(LTOD_TO_STRING(86400000000000)));      // CHECK-NEXT: LTOD#00:00:00
END_FUNCTION

(* ---- to_string_duration.st ---- *)
// RUN: %COMPILE %s && %RUN | %CHECK %s
FUNCTION main : DINT
    printf('%s$N', REF(TIME_TO_STRING(T#0ms)));              // CHECK: T#0ms
    printf('%s$N', REF(TIME_TO_STRING(T#1s500ms)));          // CHECK-NEXT: T#1s500ms
    printf('%s$N', REF(TIME_TO_STRING(T#1h1s)));              // CHECK-NEXT: T#1h1s
    printf('%s$N', REF(TIME_TO_STRING(T#1d5ms)));             // CHECK-NEXT: T#1d5ms
    printf('%s$N', REF(TIME_TO_STRING(TIME#49d17h2m47s295ms))); // CHECK-NEXT: T#49d17h2m47s295ms
    printf('%s$N', REF(LTIME_TO_STRING(LTIME#1ns)));          // CHECK-NEXT: LTIME#1ns
    printf('%s$N', REF(LTIME_TO_STRING(LTIME#1d7ns)));        // CHECK-NEXT: LTIME#1d7ns
    printf('%s$N', REF(LTIME_TO_STRING(LWORD_TO_LTIME(LWORD#18446744073709551615)))); // CHECK-NEXT: LTIME#213503d23h34m33s709ms551us615ns
    printf('%s$N', REF(TIME_TO_STRING(-1)));                  // CHECK-NEXT: T#49d17h2m47s295ms
    printf('%s$N', REF(LTIME_TO_STRING(-1)));                 // CHECK-NEXT: LTIME#213503d23h34m33s709ms551us615ns
    printf('%s$N', REF(TIME_TO_STRING(T#50d)));               // CHECK-NEXT: T#6h57m12s704ms
    printf('%s$N', REF(TIME_TO_STRING(4320000000)));          // CHECK-NEXT: T#6h57m12s704ms
    printf('%s$N', REF(LTIME_TO_STRING(9223372800000000000)));// CHECK-NEXT: LTIME#106752d
END_FUNCTION

(* ---- to_string_integer.st ---- *)
// RUN: %COMPILE %s && %RUN | %CHECK %s
FUNCTION main : DINT
    printf('%s$N', REF(BYTE_TO_STRING(BYTE#255)));       // CHECK: 255
    printf('%s$N', REF(USINT_TO_STRING(USINT#255)));     // CHECK-NEXT: 255
    printf('%s$N', REF(WORD_TO_STRING(WORD#65535)));     // CHECK-NEXT: 65535
    printf('%s$N', REF(UINT_TO_STRING(UINT#65535)));     // CHECK-NEXT: 65535
    printf('%s$N', REF(DWORD_TO_STRING(DWORD#4294967295))); // CHECK-NEXT: 4294967295
    printf('%s$N', REF(UDINT_TO_STRING(UDINT#4294967295))); // CHECK-NEXT: 4294967295
    printf('%s$N', REF(LWORD_TO_STRING(LWORD#18446744073709551615))); // CHECK-NEXT: 18446744073709551615
    printf('%s$N', REF(ULINT_TO_STRING(ULINT#18446744073709551615))); // CHECK-NEXT: 18446744073709551615
    printf('%s$N', REF(SINT_TO_STRING(SINT#-128)));      // CHECK-NEXT: -128
    printf('%s$N', REF(INT_TO_STRING(INT#-32768)));      // CHECK-NEXT: -32768
    printf('%s$N', REF(INT_TO_STRING(INT#0)));            // CHECK-NEXT: 0
    // Untyped out-of-range numeric arguments are coerced before formatting and must not panic.
    printf('%s$N', REF(BYTE_TO_STRING(256)));                 // CHECK-NEXT: 0
    printf('%s$N', REF(USINT_TO_STRING(256)));                // CHECK-NEXT: 0
    printf('%s$N', REF(WORD_TO_STRING(65536)));               // CHECK-NEXT: 0
    printf('%s$N', REF(UINT_TO_STRING(65536)));               // CHECK-NEXT: 0
    printf('%s$N', REF(DWORD_TO_STRING(4294967296)));         // CHECK-NEXT: 0
    printf('%s$N', REF(UDINT_TO_STRING(4294967296)));         // CHECK-NEXT: 0
    printf('%s$N', REF(LWORD_TO_STRING(-1)));                 // CHECK-NEXT: 18446744073709551615
    printf('%s$N', REF(ULINT_TO_STRING(-1)));                 // CHECK-NEXT: 18446744073709551615
    printf('%s$N', REF(SINT_TO_STRING(128)));                 // CHECK-NEXT: -128
    printf('%s$N', REF(INT_TO_STRING(32768)));                // CHECK-NEXT: -32768
    printf('%s$N', REF(DINT_TO_STRING(2147483648)));          // CHECK-NEXT: -2147483648
    printf('%s$N', REF(LINT_TO_STRING(1.5)));                 // CHECK-NEXT: 1
END_FUNCTION

(* ---- to_string_numeric.st ---- *)
// RUN: %COMPILE %s && %RUN | %CHECK %s
// Regression: the generic TO_STRING / TO_WSTRING must bind to the concrete per-type
// monomorphization (e.g. TO_STRING__DINT) instead of falling back to TO_STRING__STRING and
// reinterpreting the argument's bytes. DINT#-1 is a value that used to crash at runtime.
FUNCTION main : DINT
VAR
    s : STRING;
END_VAR
    s := TO_STRING(DINT#12345);          printf('%s$N', REF(s));   // CHECK: 12345
    s := TO_STRING(DINT#-1);             printf('%s$N', REF(s));   // CHECK: -1
    s := TO_STRING(LINT#-9);             printf('%s$N', REF(s));   // CHECK: -9
    s := TO_STRING(USINT#200);           printf('%s$N', REF(s));   // CHECK: 200
    s := TO_STRING(BYTE#16#FF);          printf('%s$N', REF(s));   // CHECK: 255
    s := TO_STRING(REAL#3.14);           printf('%s$N', REF(s));   // CHECK: 3.140000
    s := TO_STRING(TIME#1s500ms);        printf('%s$N', REF(s));   // CHECK: T#1s500ms

    // TO_WSTRING(DINT) binds to TO_WSTRING__DINT. printf can't print UTF-16, so compare the result
    // directly against a WSTRING literal rather than round-tripping it back through STRING.
    IF TO_WSTRING(DINT#42) = WSTRING#"42" THEN printf('ws_dint_ok$N'); END_IF   // CHECK: ws_dint_ok
END_FUNCTION

(* ---- trunc_int.st ---- *)
// RUN: %COMPILE %s && %RUN | %CHECK %s
FUNCTION main
    // REAL
    printf('%d$N', TRUNC_SINT(REAL#5.6));       // CHECK: 5
    printf('%d$N', TRUNC_USINT(REAL#5.6));      // CHECK: 5
    printf('%d$N', TRUNC_INT(REAL#5.6));        // CHECK: 5
    printf('%d$N', TRUNC_UINT(REAL#5.6));       // CHECK: 5
    printf('%d$N', TRUNC_INT(REAL#5.6));        // CHECK: 5
    printf('%d$N', TRUNC_UINT(REAL#5.6));       // CHECK: 5
    printf('%d$N', TRUNC_DINT(REAL#5.6));       // CHECK: 5
    printf('%d$N', TRUNC_UDINT(REAL#5.6));      // CHECK: 5
    printf('%d$N', TRUNC_LINT(REAL#5.6));       // CHECK: 5
    printf('%d$N', TRUNC_ULINT(REAL#5.6));      // CHECK: 5

    printf('%d$N', TRUNC_SINT(REAL#-5.6));      // CHECK: -5
    printf('%d$N', TRUNC_INT(REAL#-5.6));       // CHECK: -5
    printf('%d$N', TRUNC_DINT(REAL#-5.6));      // CHECK: -5
    printf('%d$N', TRUNC_LINT(REAL#-5.6));      // CHECK: -5

    // LREAL
    printf('%d$N', TRUNC_SINT(LREAL#5.6));       // CHECK: 5
    printf('%d$N', TRUNC_USINT(LREAL#5.6));      // CHECK: 5
    printf('%d$N', TRUNC_INT(LREAL#5.6));        // CHECK: 5
    printf('%d$N', TRUNC_UINT(LREAL#5.6));       // CHECK: 5
    printf('%d$N', TRUNC_INT(LREAL#5.6));        // CHECK: 5
    printf('%d$N', TRUNC_UINT(LREAL#5.6));       // CHECK: 5
    printf('%d$N', TRUNC_DINT(LREAL#5.6));       // CHECK: 5
    printf('%d$N', TRUNC_UDINT(LREAL#5.6));      // CHECK: 5
    printf('%d$N', TRUNC_LINT(LREAL#5.6));       // CHECK: 5
    printf('%d$N', TRUNC_ULINT(LREAL#5.6));      // CHECK: 5

    printf('%d$N', TRUNC_SINT(LREAL#-5.6));      // CHECK: -5
    printf('%d$N', TRUNC_INT(LREAL#-5.6));       // CHECK: -5
    printf('%d$N', TRUNC_DINT(LREAL#-5.6));      // CHECK: -5
    printf('%d$N', TRUNC_LINT(LREAL#-5.6));      // CHECK: -5
END_FUNCTION

(* ---- trunc_overflow.st ---- *)
// RUN: %COMPILE %s && %RUN | %CHECK %s
//
// REAL and LREAL to the integer types truncate toward zero. For SINT, USINT, INT, UINT and DINT, the
// truncated value then becomes a signed 32-bit integer and keeps the low bits of the target width;
// NaN, the infinities and anything outside the 32-bit range become -2^31, so DINT sees -2147483648
// and the narrower targets 0. UDINT, LINT and ULINT go through a signed 64-bit integer the same way
// (-2^63 when out of range), so UDINT is exact up to 2^32, and ULINT keeps a value in [2^63, 2^64)
// exact. The INT and DINT cells of the rows that the CODESYS sheet covers were measured on CODESYS
// 3.5 SP22 on x86-64 (TRUNC_INT and TRUNC, the only two truncations it provides); the other rows and
// columns extend the same rule. Each line prints SINT USINT INT UINT DINT UDINT LINT ULINT.
FUNCTION typed_real
VAR_INPUT
    x : REAL;
END_VAR
    printf('%d %d %d %d %d %u %lld %llu$N',
        REAL_TRUNC_SINT(x), REAL_TRUNC_USINT(x), REAL_TRUNC_INT(x), REAL_TRUNC_UINT(x),
        REAL_TRUNC_DINT(x), REAL_TRUNC_UDINT(x), REAL_TRUNC_LINT(x), REAL_TRUNC_ULINT(x));
END_FUNCTION

FUNCTION typed_lreal
VAR_INPUT
    x : LREAL;
END_VAR
    printf('%d %d %d %d %d %u %lld %llu$N',
        LREAL_TRUNC_SINT(x), LREAL_TRUNC_USINT(x), LREAL_TRUNC_INT(x), LREAL_TRUNC_UINT(x),
        LREAL_TRUNC_DINT(x), LREAL_TRUNC_UDINT(x), LREAL_TRUNC_LINT(x), LREAL_TRUNC_ULINT(x));
END_FUNCTION

FUNCTION generic_real
VAR_INPUT
    x : REAL;
END_VAR
    printf('%d %d %d %d %d %u %lld %llu$N',
        TRUNC_SINT(x), TRUNC_USINT(x), TRUNC_INT(x), TRUNC_UINT(x),
        TRUNC_DINT(x), TRUNC_UDINT(x), TRUNC_LINT(x), TRUNC_ULINT(x));
END_FUNCTION

FUNCTION generic_lreal
VAR_INPUT
    x : LREAL;
END_VAR
    printf('%d %d %d %d %d %u %lld %llu$N',
        TRUNC_SINT(x), TRUNC_USINT(x), TRUNC_INT(x), TRUNC_UINT(x),
        TRUNC_DINT(x), TRUNC_UDINT(x), TRUNC_LINT(x), TRUNC_ULINT(x));
END_FUNCTION

FUNCTION main
VAR
    ninf  : REAL;
    lninf : LREAL;
END_VAR
ninf  := -INF_REAL;
lninf := -INF_LREAL;

// ---- REAL source, typed form
// truncation toward zero
typed_real(REAL#5.9);       // CHECK: 5 5 5 5 5 5 5 5
typed_real(REAL#-5.9);      // CHECK: -5 251 -5 65531 -5 4294967291 -5 18446744073709551611
typed_real(REAL#-0.9);      // CHECK: 0 0 0 0 0 0 0 0
typed_real(REAL#-1.9);      // CHECK: -1 255 -1 65535 -1 4294967295 -1 18446744073709551615
// inside the 32-bit range, wraps modulo the target width
typed_real(REAL#300.7);     // CHECK: 44 44 300 300 300 300 300 300
typed_real(REAL#40000.9);   // CHECK: 64 64 -25536 40000 40000 40000 40000 40000
// outside the 32-bit range: -2^31 for SINT to DINT, while UDINT stays exact up to 2^32
typed_real(REAL#3.0E9);     // CHECK: 0 0 0 0 -2147483648 3000000000 3000000000 3000000000
typed_real(REAL#1.0E10);    // CHECK: 0 0 0 0 -2147483648 1410065408 10000000000 10000000000
typed_real(REAL#1.0E19);    // CHECK: 0 0 0 0 -2147483648 0 -9223372036854775808 9999999980506447872
typed_real(REAL#1.0E20);    // CHECK: 0 0 0 0 -2147483648 0 -9223372036854775808 9223372036854775808
// not a number
typed_real(INF_REAL);       // CHECK: 0 0 0 0 -2147483648 0 -9223372036854775808 9223372036854775808
typed_real(ninf);           // CHECK: 0 0 0 0 -2147483648 0 -9223372036854775808 9223372036854775808
typed_real(NAN_REAL);       // CHECK: 0 0 0 0 -2147483648 0 -9223372036854775808 9223372036854775808

// ---- LREAL source, typed form
typed_lreal(LREAL#-5.9);           // CHECK: -5 251 -5 65531 -5 4294967291 -5 18446744073709551611
typed_lreal(LREAL#300.7);          // CHECK: 44 44 300 300 300 300 300 300
typed_lreal(LREAL#40000.9);        // CHECK: 64 64 -25536 40000 40000 40000 40000 40000
// the edges of the 32-bit range
typed_lreal(LREAL#2147483647.9);   // CHECK: -1 255 -1 65535 2147483647 2147483647 2147483647 2147483647
typed_lreal(LREAL#2147483648.0);   // CHECK: 0 0 0 0 -2147483648 2147483648 2147483648 2147483648
typed_lreal(LREAL#-2147483648.9);  // CHECK: 0 0 0 0 -2147483648 2147483648 -2147483648 18446744071562067968
typed_lreal(LREAL#4294967295.9);   // CHECK: 0 0 0 0 -2147483648 4294967295 4294967295 4294967295
typed_lreal(LREAL#4294967296.0);   // CHECK: 0 0 0 0 -2147483648 0 4294967296 4294967296
typed_lreal(LREAL#1.0E10);         // CHECK: 0 0 0 0 -2147483648 1410065408 10000000000 10000000000
// the 64-bit band: ULINT keeps [2^63, 2^64) exact, LINT goes through the signed path
typed_lreal(LREAL#1.0E19);         // CHECK: 0 0 0 0 -2147483648 0 -9223372036854775808 10000000000000000000
typed_lreal(LREAL#-1.0E19);        // CHECK: 0 0 0 0 -2147483648 0 -9223372036854775808 9223372036854775808
typed_lreal(LREAL#1.0E20);         // CHECK: 0 0 0 0 -2147483648 0 -9223372036854775808 9223372036854775808
typed_lreal(lninf);                // CHECK: 0 0 0 0 -2147483648 0 -9223372036854775808 9223372036854775808
typed_lreal(NAN_LREAL);            // CHECK: 0 0 0 0 -2147483648 0 -9223372036854775808 9223372036854775808

// ---- the generic form calls the typed one
generic_real(REAL#-5.9);       // CHECK: -5 251 -5 65531 -5 4294967291 -5 18446744073709551611
generic_real(REAL#1.0E10);     // CHECK: 0 0 0 0 -2147483648 1410065408 10000000000 10000000000
generic_real(NAN_REAL);        // CHECK: 0 0 0 0 -2147483648 0 -9223372036854775808 9223372036854775808
generic_lreal(LREAL#40000.9);  // CHECK: 64 64 -25536 40000 40000 40000 40000 40000
generic_lreal(LREAL#1.0E19);   // CHECK: 0 0 0 0 -2147483648 0 -9223372036854775808 10000000000000000000

// ---- the deprecated TRUNC gives DINT, as TRUNC_DINT does
printf('%d %d %d %d$N', TRUNC(REAL#-5.9), TRUNC(LREAL#2147483647.9), TRUNC(LREAL#1.0E19), TRUNC(NAN_LREAL));  // CHECK: -5 2147483647 -2147483648 -2147483648
END_FUNCTION

(* ---- wstring_to_num_invalid.st ---- *)
// Malformed WSTRINGs must not crash the application; WSTRING_TO_* delegates to STRING_TO_* after a
// WSTRING->STRING conversion.

// RUN: %COMPILE %s && %RUN | %CHECK %s
FUNCTION main
    // WSTRING_TO_REAL / WSTRING_TO_LREAL: parse the valid prefix, default to 0.0
    printf('%f$N', WSTRING_TO_REAL(""));             // CHECK: 0.000000
    printf('%f$N', WSTRING_TO_REAL("asdf"));         // CHECK: 0.000000
    printf('%f$N', WSTRING_TO_REAL("1.2j3"));        // CHECK: 1.200000
    printf('%f$N', WSTRING_TO_REAL("12j3"));         // CHECK: 12.000000
    printf('%f$N', WSTRING_TO_REAL("123.456$R$N"));  // CHECK: 123.456001
    printf('%f$N', WSTRING_TO_LREAL(""));            // CHECK: 0.000000
    printf('%f$N', WSTRING_TO_LREAL("1.2j3"));       // CHECK: 1.200000

    // WSTRING_TO_DINT / WSTRING_TO_LINT: reject malformed input, default to 0
    printf('%d$N', WSTRING_TO_DINT(""));             // CHECK: 0
    printf('%d$N', WSTRING_TO_DINT("asdf"));         // CHECK: 0
    printf('%d$N', WSTRING_TO_DINT("12j3"));         // CHECK: 0
    printf('%d$N', WSTRING_TO_DINT("123.456"));      // CHECK: 123
    printf('%d$N', WSTRING_TO_LINT("12j3"));         // CHECK: 0

    // WSTRING_TO_DINT applies the DINT range, not the LINT range.
    printf('%d$N', WSTRING_TO_DINT("2147483647"));   // CHECK: 2147483647
    printf('%d$N', WSTRING_TO_DINT("2147483648"));   // CHECK: 0
    printf('%d$N', WSTRING_TO_DINT("4294967297"));   // CHECK: 0
END_FUNCTION

(* ---- bool_constant_values.st ---- *)
// RUN: not %COMPILE --error-format clang %s 2>&1 | %CHECK --implicit-check-not='{{.*}}error[E037]{{.*}}' %s

// A constant integer value other than 0 or 1 is no BOOL value. The compiler rejects it in a
// body assignment, an initializer and a call argument, whatever form computes the value.
// The values 0 and 1, non-constant integers, and members whose name matches a constant stay valid.

TYPE State : (idle, running, done); END_TYPE

VAR_GLOBAL CONSTANT
    cTwo : INT := 2;
    cOne : INT := 1;
    cFalse : BOOL := 0;
END_VAR

FUNCTION takesBool : BOOL
VAR_INPUT
    x : BOOL;
END_VAR
    takesBool := x;
END_FUNCTION

FUNCTION_BLOCK withProperty
VAR
    _p : BOOL;
END_VAR
PROPERTY_SET prop : BOOL
    _p := prop;
END_PROPERTY
END_FUNCTION_BLOCK

FUNCTION_BLOCK Base
VAR_OUTPUT
    done : BOOL;
END_VAR
END_FUNCTION_BLOCK

FUNCTION_BLOCK Derived EXTENDS Base
VAR
    last : BOOL;
END_VAR
    last := done;
    last := SUPER^.done;
END_FUNCTION_BLOCK

PROGRAM mainProg
VAR
    inst : withProperty;
    // CHECK-DAG: {{.*}}bool_constant_values.st:[[@LINE+1]]:{{[0-9]+}}:{{.*}}error[E037]: Invalid assignment: cannot assign the value 2 to 'BOOL'
    fromConstant : BOOL := cTwo;
    validFromConstant : BOOL := cOne;
    b : BOOL;
    i : DINT;
    d : Derived;
END_VAR
    // CHECK-DAG: {{.*}}bool_constant_values.st:[[@LINE+1]]:{{[0-9]+}}:{{.*}}error[E037]: Invalid assignment: cannot assign the value 5 to 'BOOL'
    b := INT#5;
    // CHECK-DAG: {{.*}}bool_constant_values.st:[[@LINE+1]]:{{[0-9]+}}:{{.*}}error[E037]: Invalid assignment: cannot assign the value 2 to 'BOOL'
    b := 1 + 1;
    // CHECK-DAG: {{.*}}bool_constant_values.st:[[@LINE+1]]:{{[0-9]+}}:{{.*}}error[E037]: Invalid assignment: cannot assign the value 3 to 'BOOL'
    takesBool(INT#3);
    // CHECK-DAG: {{.*}}bool_constant_values.st:[[@LINE+1]]:{{[0-9]+}}:{{.*}}error[E037]: Invalid assignment: cannot assign the value 4 to 'BOOL'
    inst.prop := INT#4;
    inst.prop := INT#1;
    b := INT#1;
    b := 1 * 1;
    b := i;
    takesBool(cOne);
    b := d.done;
    b := NOT cFalse;
END_PROGRAM
